(* IEC 61131-3 sources: deprecated-refusr-repo/samples (part 8) *)

(* ---- 4-MUX_golem-sudsy-awing.st ---- *)
(*
This code implements a shuffled multiplexer with 4 control bits.
The control bits are: Data[N2], Data[N3], Data[N4], Data[N6]
The input bits are: Data[N1], Data[N5], Data[N8], Data[N9], Data[N7], Data[N12], Data[N10], Data[N17], Data[N11], Data[N18], Data[N14], Data[N13], Data[N20], Data[N15], Data[N16], Data[N19]

The symbolic expression is:
((((((((((((((((!((((!(IN2)) & (!(IN3))) & (!(IN4))) & (!(IN6)))) | IN1) & ((!(((IN2 & (!(IN3))) & (!(IN4))) & (!(IN6)))) | IN5)) & ((!((((!(IN2)) & IN3) & (!(IN4))) & (!(IN6)))) | IN8)) & ((!(((IN2 & IN3) & (!(IN4))) & (!(IN6)))) | IN9)) & ((!((((!(IN2)) & (!(IN3))) & IN4) & (!(IN6)))) | IN7)) & ((!(((IN2 & (!(IN3))) & IN4) & (!(IN6)))) | IN12)) & ((!((((!(IN2)) & IN3) & IN4) & (!(IN6)))) | IN10)) & ((!(((IN2 & IN3) & IN4) & (!(IN6)))) | IN17)) & ((!((((!(IN2)) & (!(IN3))) & (!(IN4))) & IN6)) | IN11)) & ((!(((IN2 & (!(IN3))) & (!(IN4))) & IN6)) | IN18)) & ((!((((!(IN2)) & IN3) & (!(IN4))) & IN6)) | IN14)) & ((!(((IN2 & IN3) & (!(IN4))) & IN6)) | IN13)) & ((!((((!(IN2)) & (!(IN3))) & IN4) & IN6)) | IN20)) & ((!(((IN2 & (!(IN3))) & IN4) & IN6)) | IN15)) & ((!((((!(IN2)) & IN3) & IN4) & IN6)) | IN16)) & ((!(((IN2 & IN3) & IN4) & IN6)) | IN19)

*)

FUNCTION_BLOCK F_CollectInput
  VAR_IN_OUT
      Data : ARRAY[1..20] OF BOOL;
  END_VAR
  VAR_INPUT
      TICK  : BOOL := 0;
      IN1   : BOOL := 0;
      IN2   : BOOL := 0;
      IN3   : BOOL := 0;
      IN4   : BOOL := 0;
      IN5   : BOOL := 0;
      RESET : BOOL := FALSE;
  END_VAR
  VAR_OUTPUT
      Finished : BOOL;
  END_VAR
  VAR
      j    : USINT := 1;
      tock : BOOL  := 0;
  END_VAR
  IF NOT RESET AND tock = NOT TICK THEN
      Data[j]   := IN1;
      Data[j+1] := IN2;
      Data[j+2] := IN3;
      Data[j+3] := IN4;
      Data[j+4] := IN5;
      j := j + 5;
      tock := TICK;
  ELSE
      j := 1;
      tock := 0;
  END_IF;
  Finished := (j > 20);
END_FUNCTION_BLOCK

PROGRAM Boiler
  VAR
    Data  : ARRAY[1..20] OF BOOL;
    Ready : BOOL;
    CollectInput : F_CollectInput;
  END_VAR
  VAR
    TICK     AT %IX1.0 : BOOL;
    IN1      AT %IX0.3 : BOOL;
    IN2      AT %IX0.4 : BOOL;
    IN3      AT %IX0.5 : BOOL;
    IN4      AT %IX0.6 : BOOL;
    IN5      AT %IX0.7 : BOOL;
    OutReady AT %QX0.0 : BOOL := FALSE;
    FeedNext AT %QX0.1 : BOOL := FALSE;
    Out      AT %QX0.2 : BOOL;
  END_VAR
  CollectInput(TICK:=TICK, IN1:=IN1, IN2:=IN2, IN3:=IN3, IN4:=IN4, IN5:=IN5);
  Ready := CollectInput.Finished;
  FeedNext := 1;
  IF Ready THEN
    Out := (((((((((((((((((NOT ((((NOT Data[2]) AND (NOT Data[3])) AND (NOT Data[4])) AND (NOT Data[6]))) OR Data[1]) AND ((NOT (((Data[2] AND (NOT Data[3])) AND (NOT Data[4])) AND (NOT Data[6]))) OR Data[5])) AND ((NOT ((((NOT Data[2]) AND Data[3]) AND (NOT Data[4])) AND (NOT Data[6]))) OR Data[8])) AND ((NOT (((Data[2] AND Data[3]) AND (NOT Data[4])) AND (NOT Data[6]))) OR Data[9])) AND ((NOT ((((NOT Data[2]) AND (NOT Data[3])) AND Data[4]) AND (NOT Data[6]))) OR Data[7])) AND ((NOT (((Data[2] AND (NOT Data[3])) AND Data[4]) AND (NOT Data[6]))) OR Data[12])) AND ((NOT ((((NOT Data[2]) AND Data[3]) AND Data[4]) AND (NOT Data[6]))) OR Data[10])) AND ((NOT (((Data[2] AND Data[3]) AND Data[4]) AND (NOT Data[6]))) OR Data[17])) AND ((NOT ((((NOT Data[2]) AND (NOT Data[3])) AND (NOT Data[4])) AND Data[6])) OR Data[11])) AND ((NOT (((Data[2] AND (NOT Data[3])) AND (NOT Data[4])) AND Data[6])) OR Data[18])) AND ((NOT ((((NOT Data[2]) AND Data[3]) AND (NOT Data[4])) AND Data[6])) OR Data[14])) AND ((NOT (((Data[2] AND Data[3]) AND (NOT Data[4])) AND Data[6])) OR Data[13])) AND ((NOT ((((NOT Data[2]) AND (NOT Data[3])) AND Data[4]) AND Data[6])) OR Data[20])) AND ((NOT (((Data[2] AND (NOT Data[3])) AND Data[4]) AND Data[6])) OR Data[15])) AND ((NOT ((((NOT Data[2]) AND Data[3]) AND Data[4]) AND Data[6])) OR Data[16])) AND ((NOT (((Data[2] AND Data[3]) AND Data[4]) AND Data[6])) OR Data[19]));
    OutReady := 1;
    CollectInput(RESET:=TRUE);
  END_IF;
END_PROGRAM

CONFIGURATION Config0
  RESOURCE Res0 ON PLC
    TASK task0(INTERVAL := T#20ms,PRIORITY := 0);
    PROGRAM instance0 WITH task0 : Boiler;
  END_RESOURCE
END_CONFIGURATION

(* ---- 4-MUX_grout-chafe-snail.st ---- *)
(*
This code implements a shuffled multiplexer with 4 control bits.
The control bits are: Data[N8], Data[N2], Data[N5], Data[N1]
The input bits are: Data[N4], Data[N11], Data[N3], Data[N7], Data[N6], Data[N9], Data[N14], Data[N12], Data[N13], Data[N15], Data[N16], Data[N17], Data[N19], Data[N20], Data[N10], Data[N18]

The symbolic expression is:
((((((((((((((((!((((!(IN8)) & (!(IN2))) & (!(IN5))) & (!(IN1)))) | IN4) & ((!(((IN8 & (!(IN2))) & (!(IN5))) & (!(IN1)))) | IN11)) & ((!((((!(IN8)) & IN2) & (!(IN5))) & (!(IN1)))) | IN3)) & ((!(((IN8 & IN2) & (!(IN5))) & (!(IN1)))) | IN7)) & ((!((((!(IN8)) & (!(IN2))) & IN5) & (!(IN1)))) | IN6)) & ((!(((IN8 & (!(IN2))) & IN5) & (!(IN1)))) | IN9)) & ((!((((!(IN8)) & IN2) & IN5) & (!(IN1)))) | IN14)) & ((!(((IN8 & IN2) & IN5) & (!(IN1)))) | IN12)) & ((!((((!(IN8)) & (!(IN2))) & (!(IN5))) & IN1)) | IN13)) & ((!(((IN8 & (!(IN2))) & (!(IN5))) & IN1)) | IN15)) & ((!((((!(IN8)) & IN2) & (!(IN5))) & IN1)) | IN16)) & ((!(((IN8 & IN2) & (!(IN5))) & IN1)) | IN17)) & ((!((((!(IN8)) & (!(IN2))) & IN5) & IN1)) | IN19)) & ((!(((IN8 & (!(IN2))) & IN5) & IN1)) | IN20)) & ((!((((!(IN8)) & IN2) & IN5) & IN1)) | IN10)) & ((!(((IN8 & IN2) & IN5) & IN1)) | IN18)

*)

FUNCTION_BLOCK F_CollectInput
  VAR_IN_OUT
      Data : ARRAY[1..20] OF BOOL;
  END_VAR
  VAR_INPUT
      TICK  : BOOL := 0;
      IN1   : BOOL := 0;
      IN2   : BOOL := 0;
      IN3   : BOOL := 0;
      IN4   : BOOL := 0;
      IN5   : BOOL := 0;
      RESET : BOOL := FALSE;
  END_VAR
  VAR_OUTPUT
      Finished : BOOL;
  END_VAR
  VAR
      j    : USINT := 1;
      tock : BOOL  := 0;
  END_VAR
  IF NOT RESET AND tock = NOT TICK THEN
      Data[j]   := IN1;
      Data[j+1] := IN2;
      Data[j+2] := IN3;
      Data[j+3] := IN4;
      Data[j+4] := IN5;
      j := j + 5;
      tock := TICK;
  ELSE
      j := 1;
      tock := 0;
  END_IF;
  Finished := (j > 20);
END_FUNCTION_BLOCK

PROGRAM Boiler
  VAR
    Data  : ARRAY[1..20] OF BOOL;
    Ready : BOOL;
    CollectInput : F_CollectInput;
  END_VAR
  VAR
    TICK     AT %IX1.0 : BOOL;
    IN1      AT %IX0.3 : BOOL;
    IN2      AT %IX0.4 : BOOL;
    IN3      AT %IX0.5 : BOOL;
    IN4      AT %IX0.6 : BOOL;
    IN5      AT %IX0.7 : BOOL;
    OutReady AT %QX0.0 : BOOL := FALSE;
    FeedNext AT %QX0.1 : BOOL := FALSE;
    Out      AT %QX0.2 : BOOL;
  END_VAR
  CollectInput(TICK:=TICK, IN1:=IN1, IN2:=IN2, IN3:=IN3, IN4:=IN4, IN5:=IN5);
  Ready := CollectInput.Finished;
  FeedNext := 1;
  IF Ready THEN
    Out := (((((((((((((((((NOT ((((NOT Data[8]) AND (NOT Data[2])) AND (NOT Data[5])) AND (NOT Data[1]))) OR Data[4]) AND ((NOT (((Data[8] AND (NOT Data[2])) AND (NOT Data[5])) AND (NOT Data[1]))) OR Data[11])) AND ((NOT ((((NOT Data[8]) AND Data[2]) AND (NOT Data[5])) AND (NOT Data[1]))) OR Data[3])) AND ((NOT (((Data[8] AND Data[2]) AND (NOT Data[5])) AND (NOT Data[1]))) OR Data[7])) AND ((NOT ((((NOT Data[8]) AND (NOT Data[2])) AND Data[5]) AND (NOT Data[1]))) OR Data[6])) AND ((NOT (((Data[8] AND (NOT Data[2])) AND Data[5]) AND (NOT Data[1]))) OR Data[9])) AND ((NOT ((((NOT Data[8]) AND Data[2]) AND Data[5]) AND (NOT Data[1]))) OR Data[14])) AND ((NOT (((Data[8] AND Data[2]) AND Data[5]) AND (NOT Data[1]))) OR Data[12])) AND ((NOT ((((NOT Data[8]) AND (NOT Data[2])) AND (NOT Data[5])) AND Data[1])) OR Data[13])) AND ((NOT (((Data[8] AND (NOT Data[2])) AND (NOT Data[5])) AND Data[1])) OR Data[15])) AND ((NOT ((((NOT Data[8]) AND Data[2]) AND (NOT Data[5])) AND Data[1])) OR Data[16])) AND ((NOT (((Data[8] AND Data[2]) AND (NOT Data[5])) AND Data[1])) OR Data[17])) AND ((NOT ((((NOT Data[8]) AND (NOT Data[2])) AND Data[5]) AND Data[1])) OR Data[19])) AND ((NOT (((Data[8] AND (NOT Data[2])) AND Data[5]) AND Data[1])) OR Data[20])) AND ((NOT ((((NOT Data[8]) AND Data[2]) AND Data[5]) AND Data[1])) OR Data[10])) AND ((NOT (((Data[8] AND Data[2]) AND Data[5]) AND Data[1])) OR Data[18]));
    OutReady := 1;
    CollectInput(RESET:=TRUE);
  END_IF;
END_PROGRAM

CONFIGURATION Config0
  RESOURCE Res0 ON PLC
    TASK task0(INTERVAL := T#20ms,PRIORITY := 0);
    PROGRAM instance0 WITH task0 : Boiler;
  END_RESOURCE
END_CONFIGURATION

(* ---- 4-MUX_grump-gavel-russe.st ---- *)
(*
This code implements a shuffled multiplexer with 4 control bits.
The control bits are: Data[N2], Data[N3], Data[N4], Data[N7]
The input bits are: Data[N1], Data[N5], Data[N10], Data[N6], Data[N8], Data[N9], Data[N12], Data[N13], Data[N11], Data[N14], Data[N15], Data[N16], Data[N17], Data[N18], Data[N19], Data[N20]

The symbolic expression is:
((((((((((((((((!((((!(IN2)) & (!(IN3))) & (!(IN4))) & (!(IN7)))) | IN1) & ((!(((IN2 & (!(IN3))) & (!(IN4))) & (!(IN7)))) | IN5)) & ((!((((!(IN2)) & IN3) & (!(IN4))) & (!(IN7)))) | IN10)) & ((!(((IN2 & IN3) & (!(IN4))) & (!(IN7)))) | IN6)) & ((!((((!(IN2)) & (!(IN3))) & IN4) & (!(IN7)))) | IN8)) & ((!(((IN2 & (!(IN3))) & IN4) & (!(IN7)))) | IN9)) & ((!((((!(IN2)) & IN3) & IN4) & (!(IN7)))) | IN12)) & ((!(((IN2 & IN3) & IN4) & (!(IN7)))) | IN13)) & ((!((((!(IN2)) & (!(IN3))) & (!(IN4))) & IN7)) | IN11)) & ((!(((IN2 & (!(IN3))) & (!(IN4))) & IN7)) | IN14)) & ((!((((!(IN2)) & IN3) & (!(IN4))) & IN7)) | IN15)) & ((!(((IN2 & IN3) & (!(IN4))) & IN7)) | IN16)) & ((!((((!(IN2)) & (!(IN3))) & IN4) & IN7)) | IN17)) & ((!(((IN2 & (!(IN3))) & IN4) & IN7)) | IN18)) & ((!((((!(IN2)) & IN3) & IN4) & IN7)) | IN19)) & ((!(((IN2 & IN3) & IN4) & IN7)) | IN20)

*)

FUNCTION_BLOCK F_CollectInput
  VAR_IN_OUT
      Data : ARRAY[1..20] OF BOOL;
  END_VAR
  VAR_INPUT
      TICK  : BOOL := 0;
      IN1   : BOOL := 0;
      IN2   : BOOL := 0;
      IN3   : BOOL := 0;
      IN4   : BOOL := 0;
      IN5   : BOOL := 0;
      RESET : BOOL := FALSE;
  END_VAR
  VAR_OUTPUT
      Finished : BOOL;
  END_VAR
  VAR
      j    : USINT := 1;
      tock : BOOL  := 0;
  END_VAR
  IF NOT RESET AND tock = NOT TICK THEN
      Data[j]   := IN1;
      Data[j+1] := IN2;
      Data[j+2] := IN3;
      Data[j+3] := IN4;
      Data[j+4] := IN5;
      j := j + 5;
      tock := TICK;
  ELSE
      j := 1;
      tock := 0;
  END_IF;
  Finished := (j > 20);
END_FUNCTION_BLOCK

PROGRAM Boiler
  VAR
    Data  : ARRAY[1..20] OF BOOL;
    Ready : BOOL;
    CollectInput : F_CollectInput;
  END_VAR
  VAR
    TICK     AT %IX1.0 : BOOL;
    IN1      AT %IX0.3 : BOOL;
    IN2      AT %IX0.4 : BOOL;
    IN3      AT %IX0.5 : BOOL;
    IN4      AT %IX0.6 : BOOL;
    IN5      AT %IX0.7 : BOOL;
    OutReady AT %QX0.0 : BOOL := FALSE;
    FeedNext AT %QX0.1 : BOOL := FALSE;
    Out      AT %QX0.2 : BOOL;
  END_VAR
  CollectInput(TICK:=TICK, IN1:=IN1, IN2:=IN2, IN3:=IN3, IN4:=IN4, IN5:=IN5);
  Ready := CollectInput.Finished;
  FeedNext := 1;
  IF Ready THEN
    Out := (((((((((((((((((NOT ((((NOT Data[2]) AND (NOT Data[3])) AND (NOT Data[4])) AND (NOT Data[7]))) OR Data[1]) AND ((NOT (((Data[2] AND (NOT Data[3])) AND (NOT Data[4])) AND (NOT Data[7]))) OR Data[5])) AND ((NOT ((((NOT Data[2]) AND Data[3]) AND (NOT Data[4])) AND (NOT Data[7]))) OR Data[10])) AND ((NOT (((Data[2] AND Data[3]) AND (NOT Data[4])) AND (NOT Data[7]))) OR Data[6])) AND ((NOT ((((NOT Data[2]) AND (NOT Data[3])) AND Data[4]) AND (NOT Data[7]))) OR Data[8])) AND ((NOT (((Data[2] AND (NOT Data[3])) AND Data[4]) AND (NOT Data[7]))) OR Data[9])) AND ((NOT ((((NOT Data[2]) AND Data[3]) AND Data[4]) AND (NOT Data[7]))) OR Data[12])) AND ((NOT (((Data[2] AND Data[3]) AND Data[4]) AND (NOT Data[7]))) OR Data[13])) AND ((NOT ((((NOT Data[2]) AND (NOT Data[3])) AND (NOT Data[4])) AND Data[7])) OR Data[11])) AND ((NOT (((Data[2] AND (NOT Data[3])) AND (NOT Data[4])) AND Data[7])) OR Data[14])) AND ((NOT ((((NOT Data[2]) AND Data[3]) AND (NOT Data[4])) AND Data[7])) OR Data[15])) AND ((NOT (((Data[2] AND Data[3]) AND (NOT Data[4])) AND Data[7])) OR Data[16])) AND ((NOT ((((NOT Data[2]) AND (NOT Data[3])) AND Data[4]) AND Data[7])) OR Data[17])) AND ((NOT (((Data[2] AND (NOT Data[3])) AND Data[4]) AND Data[7])) OR Data[18])) AND ((NOT ((((NOT Data[2]) AND Data[3]) AND Data[4]) AND Data[7])) OR Data[19])) AND ((NOT (((Data[2] AND Data[3]) AND Data[4]) AND Data[7])) OR Data[20]));
    OutReady := 1;
    CollectInput(RESET:=TRUE);
  END_IF;
END_PROGRAM

CONFIGURATION Config0
  RESOURCE Res0 ON PLC
    TASK task0(INTERVAL := T#20ms,PRIORITY := 0);
    PROGRAM instance0 WITH task0 : Boiler;
  END_RESOURCE
END_CONFIGURATION

(* ---- 4-MUX_gyved-gauzy-steed.st ---- *)
(*
This code implements a shuffled multiplexer with 4 control bits.
The control bits are: Data[N3], Data[N4], Data[N1], Data[N6]
The input bits are: Data[N2], Data[N10], Data[N9], Data[N5], Data[N7], Data[N11], Data[N8], Data[N12], Data[N14], Data[N13], Data[N15], Data[N18], Data[N16], Data[N17], Data[N19], Data[N20]

The symbolic expression is:
((((((((((((((((!((((!(IN3)) & (!(IN4))) & (!(IN1))) & (!(IN6)))) | IN2) & ((!(((IN3 & (!(IN4))) & (!(IN1))) & (!(IN6)))) | IN10)) & ((!((((!(IN3)) & IN4) & (!(IN1))) & (!(IN6)))) | IN9)) & ((!(((IN3 & IN4) & (!(IN1))) & (!(IN6)))) | IN5)) & ((!((((!(IN3)) & (!(IN4))) & IN1) & (!(IN6)))) | IN7)) & ((!(((IN3 & (!(IN4))) & IN1) & (!(IN6)))) | IN11)) & ((!((((!(IN3)) & IN4) & IN1) & (!(IN6)))) | IN8)) & ((!(((IN3 & IN4) & IN1) & (!(IN6)))) | IN12)) & ((!((((!(IN3)) & (!(IN4))) & (!(IN1))) & IN6)) | IN14)) & ((!(((IN3 & (!(IN4))) & (!(IN1))) & IN6)) | IN13)) & ((!((((!(IN3)) & IN4) & (!(IN1))) & IN6)) | IN15)) & ((!(((IN3 & IN4) & (!(IN1))) & IN6)) | IN18)) & ((!((((!(IN3)) & (!(IN4))) & IN1) & IN6)) | IN16)) & ((!(((IN3 & (!(IN4))) & IN1) & IN6)) | IN17)) & ((!((((!(IN3)) & IN4) & IN1) & IN6)) | IN19)) & ((!(((IN3 & IN4) & IN1) & IN6)) | IN20)

*)

FUNCTION_BLOCK F_CollectInput
  VAR_IN_OUT
      Data : ARRAY[1..20] OF BOOL;
  END_VAR
  VAR_INPUT
      TICK  : BOOL := 0;
      IN1   : BOOL := 0;
      IN2   : BOOL := 0;
      IN3   : BOOL := 0;
      IN4   : BOOL := 0;
      IN5   : BOOL := 0;
      RESET : BOOL := FALSE;
  END_VAR
  VAR_OUTPUT
      Finished : BOOL;
  END_VAR
  VAR
      j    : USINT := 1;
      tock : BOOL  := 0;
  END_VAR
  IF NOT RESET AND tock = NOT TICK THEN
      Data[j]   := IN1;
      Data[j+1] := IN2;
      Data[j+2] := IN3;
      Data[j+3] := IN4;
      Data[j+4] := IN5;
      j := j + 5;
      tock := TICK;
  ELSE
      j := 1;
      tock := 0;
  END_IF;
  Finished := (j > 20);
END_FUNCTION_BLOCK

PROGRAM Boiler
  VAR
    Data  : ARRAY[1..20] OF BOOL;
    Ready : BOOL;
    CollectInput : F_CollectInput;
  END_VAR
  VAR
    TICK     AT %IX1.0 : BOOL;
    IN1      AT %IX0.3 : BOOL;
    IN2      AT %IX0.4 : BOOL;
    IN3      AT %IX0.5 : BOOL;
    IN4      AT %IX0.6 : BOOL;
    IN5      AT %IX0.7 : BOOL;
    OutReady AT %QX0.0 : BOOL := FALSE;
    FeedNext AT %QX0.1 : BOOL := FALSE;
    Out      AT %QX0.2 : BOOL;
  END_VAR
  CollectInput(TICK:=TICK, IN1:=IN1, IN2:=IN2, IN3:=IN3, IN4:=IN4, IN5:=IN5);
  Ready := CollectInput.Finished;
  FeedNext := 1;
  IF Ready THEN
    Out := (((((((((((((((((NOT ((((NOT Data[3]) AND (NOT Data[4])) AND (NOT Data[1])) AND (NOT Data[6]))) OR Data[2]) AND ((NOT (((Data[3] AND (NOT Data[4])) AND (NOT Data[1])) AND (NOT Data[6]))) OR Data[10])) AND ((NOT ((((NOT Data[3]) AND Data[4]) AND (NOT Data[1])) AND (NOT Data[6]))) OR Data[9])) AND ((NOT (((Data[3] AND Data[4]) AND (NOT Data[1])) AND (NOT Data[6]))) OR Data[5])) AND ((NOT ((((NOT Data[3]) AND (NOT Data[4])) AND Data[1]) AND (NOT Data[6]))) OR Data[7])) AND ((NOT (((Data[3] AND (NOT Data[4])) AND Data[1]) AND (NOT Data[6]))) OR Data[11])) AND ((NOT ((((NOT Data[3]) AND Data[4]) AND Data[1]) AND (NOT Data[6]))) OR Data[8])) AND ((NOT (((Data[3] AND Data[4]) AND Data[1]) AND (NOT Data[6]))) OR Data[12])) AND ((NOT ((((NOT Data[3]) AND (NOT Data[4])) AND (NOT Data[1])) AND Data[6])) OR Data[14])) AND ((NOT (((Data[3] AND (NOT Data[4])) AND (NOT Data[1])) AND Data[6])) OR Data[13])) AND ((NOT ((((NOT Data[3]) AND Data[4]) AND (NOT Data[1])) AND Data[6])) OR Data[15])) AND ((NOT (((Data[3] AND Data[4]) AND (NOT Data[1])) AND Data[6])) OR Data[18])) AND ((NOT ((((NOT Data[3]) AND (NOT Data[4])) AND Data[1]) AND Data[6])) OR Data[16])) AND ((NOT (((Data[3] AND (NOT Data[4])) AND Data[1]) AND Data[6])) OR Data[17])) AND ((NOT ((((NOT Data[3]) AND Data[4]) AND Data[1]) AND Data[6])) OR Data[19])) AND ((NOT (((Data[3] AND Data[4]) AND Data[1]) AND Data[6])) OR Data[20]));
    OutReady := 1;
    CollectInput(RESET:=TRUE);
  END_IF;
END_PROGRAM

CONFIGURATION Config0
  RESOURCE Res0 ON PLC
    TASK task0(INTERVAL := T#20ms,PRIORITY := 0);
    PROGRAM instance0 WITH task0 : Boiler;
  END_RESOURCE
END_CONFIGURATION

(* ---- 4-MUX_havoc-schmo-linty.st ---- *)
(*
This code implements a shuffled multiplexer with 4 control bits.
The control bits are: Data[N3], Data[N8], Data[N5], Data[N2]
The input bits are: Data[N1], Data[N9], Data[N4], Data[N6], Data[N7], Data[N10], Data[N12], Data[N11], Data[N14], Data[N13], Data[N16], Data[N15], Data[N18], Data[N19], Data[N20], Data[N17]

The symbolic expression is:
((((((((((((((((!((((!(IN3)) & (!(IN8))) & (!(IN5))) & (!(IN2)))) | IN1) & ((!(((IN3 & (!(IN8))) & (!(IN5))) & (!(IN2)))) | IN9)) & ((!((((!(IN3)) & IN8) & (!(IN5))) & (!(IN2)))) | IN4)) & ((!(((IN3 & IN8) & (!(IN5))) & (!(IN2)))) | IN6)) & ((!((((!(IN3)) & (!(IN8))) & IN5) & (!(IN2)))) | IN7)) & ((!(((IN3 & (!(IN8))) & IN5) & (!(IN2)))) | IN10)) & ((!((((!(IN3)) & IN8) & IN5) & (!(IN2)))) | IN12)) & ((!(((IN3 & IN8) & IN5) & (!(IN2)))) | IN11)) & ((!((((!(IN3)) & (!(IN8))) & (!(IN5))) & IN2)) | IN14)) & ((!(((IN3 & (!(IN8))) & (!(IN5))) & IN2)) | IN13)) & ((!((((!(IN3)) & IN8) & (!(IN5))) & IN2)) | IN16)) & ((!(((IN3 & IN8) & (!(IN5))) & IN2)) | IN15)) & ((!((((!(IN3)) & (!(IN8))) & IN5) & IN2)) | IN18)) & ((!(((IN3 & (!(IN8))) & IN5) & IN2)) | IN19)) & ((!((((!(IN3)) & IN8) & IN5) & IN2)) | IN20)) & ((!(((IN3 & IN8) & IN5) & IN2)) | IN17)

*)

FUNCTION_BLOCK F_CollectInput
  VAR_IN_OUT
      Data : ARRAY[1..20] OF BOOL;
  END_VAR
  VAR_INPUT
      TICK  : BOOL := 0;
      IN1   : BOOL := 0;
      IN2   : BOOL := 0;
      IN3   : BOOL := 0;
      IN4   : BOOL := 0;
      IN5   : BOOL := 0;
      RESET : BOOL := FALSE;
  END_VAR
  VAR_OUTPUT
      Finished : BOOL;
  END_VAR
  VAR
      j    : USINT := 1;
      tock : BOOL  := 0;
  END_VAR
  IF NOT RESET AND tock = NOT TICK THEN
      Data[j]   := IN1;
      Data[j+1] := IN2;
      Data[j+2] := IN3;
      Data[j+3] := IN4;
      Data[j+4] := IN5;
      j := j + 5;
      tock := TICK;
  ELSE
      j := 1;
      tock := 0;
  END_IF;
  Finished := (j > 20);
END_FUNCTION_BLOCK

PROGRAM Boiler
  VAR
    Data  : ARRAY[1..20] OF BOOL;
    Ready : BOOL;
    CollectInput : F_CollectInput;
  END_VAR
  VAR
    TICK     AT %IX1.0 : BOOL;
    IN1      AT %IX0.3 : BOOL;
    IN2      AT %IX0.4 : BOOL;
    IN3      AT %IX0.5 : BOOL;
    IN4      AT %IX0.6 : BOOL;
    IN5      AT %IX0.7 : BOOL;
    OutReady AT %QX0.0 : BOOL := FALSE;
    FeedNext AT %QX0.1 : BOOL := FALSE;
    Out      AT %QX0.2 : BOOL;
  END_VAR
  CollectInput(TICK:=TICK, IN1:=IN1, IN2:=IN2, IN3:=IN3, IN4:=IN4, IN5:=IN5);
  Ready := CollectInput.Finished;
  FeedNext := 1;
  IF Ready THEN
    Out := (((((((((((((((((NOT ((((NOT Data[3]) AND (NOT Data[8])) AND (NOT Data[5])) AND (NOT Data[2]))) OR Data[1]) AND ((NOT (((Data[3] AND (NOT Data[8])) AND (NOT Data[5])) AND (NOT Data[2]))) OR Data[9])) AND ((NOT ((((NOT Data[3]) AND Data[8]) AND (NOT Data[5])) AND (NOT Data[2]))) OR Data[4])) AND ((NOT (((Data[3] AND Data[8]) AND (NOT Data[5])) AND (NOT Data[2]))) OR Data[6])) AND ((NOT ((((NOT Data[3]) AND (NOT Data[8])) AND Data[5]) AND (NOT Data[2]))) OR Data[7])) AND ((NOT (((Data[3] AND (NOT Data[8])) AND Data[5]) AND (NOT Data[2]))) OR Data[10])) AND ((NOT ((((NOT Data[3]) AND Data[8]) AND Data[5]) AND (NOT Data[2]))) OR Data[12])) AND ((NOT (((Data[3] AND Data[8]) AND Data[5]) AND (NOT Data[2]))) OR Data[11])) AND ((NOT ((((NOT Data[3]) AND (NOT Data[8])) AND (NOT Data[5])) AND Data[2])) OR Data[14])) AND ((NOT (((Data[3] AND (NOT Data[8])) AND (NOT Data[5])) AND Data[2])) OR Data[13])) AND ((NOT ((((NOT Data[3]) AND Data[8]) AND (NOT Data[5])) AND Data[2])) OR Data[16])) AND ((NOT (((Data[3] AND Data[8]) AND (NOT Data[5])) AND Data[2])) OR Data[15])) AND ((NOT ((((NOT Data[3]) AND (NOT Data[8])) AND Data[5]) AND Data[2])) OR Data[18])) AND ((NOT (((Data[3] AND (NOT Data[8])) AND Data[5]) AND Data[2])) OR Data[19])) AND ((NOT ((((NOT Data[3]) AND Data[8]) AND Data[5]) AND Data[2])) OR Data[20])) AND ((NOT (((Data[3] AND Data[8]) AND Data[5]) AND Data[2])) OR Data[17]));
    OutReady := 1;
    CollectInput(RESET:=TRUE);
  END_IF;
END_PROGRAM

CONFIGURATION Config0
  RESOURCE Res0 ON PLC
    TASK task0(INTERVAL := T#20ms,PRIORITY := 0);
    PROGRAM instance0 WITH task0 : Boiler;
  END_RESOURCE
END_CONFIGURATION

(* ---- 4-MUX_holds-splat-brent.st ---- *)
(*
This code implements a shuffled multiplexer with 4 control bits.
The control bits are: Data[N1], Data[N4], Data[N5], Data[N3]
The input bits are: Data[N2], Data[N7], Data[N11], Data[N6], Data[N8], Data[N12], Data[N9], Data[N10], Data[N16], Data[N14], Data[N13], Data[N18], Data[N17], Data[N15], Data[N19], Data[N20]

The symbolic expression is:
((((((((((((((((!((((!(IN1)) & (!(IN4))) & (!(IN5))) & (!(IN3)))) | IN2) & ((!(((IN1 & (!(IN4))) & (!(IN5))) & (!(IN3)))) | IN7)) & ((!((((!(IN1)) & IN4) & (!(IN5))) & (!(IN3)))) | IN11)) & ((!(((IN1 & IN4) & (!(IN5))) & (!(IN3)))) | IN6)) & ((!((((!(IN1)) & (!(IN4))) & IN5) & (!(IN3)))) | IN8)) & ((!(((IN1 & (!(IN4))) & IN5) & (!(IN3)))) | IN12)) & ((!((((!(IN1)) & IN4) & IN5) & (!(IN3)))) | IN9)) & ((!(((IN1 & IN4) & IN5) & (!(IN3)))) | IN10)) & ((!((((!(IN1)) & (!(IN4))) & (!(IN5))) & IN3)) | IN16)) & ((!(((IN1 & (!(IN4))) & (!(IN5))) & IN3)) | IN14)) & ((!((((!(IN1)) & IN4) & (!(IN5))) & IN3)) | IN13)) & ((!(((IN1 & IN4) & (!(IN5))) & IN3)) | IN18)) & ((!((((!(IN1)) & (!(IN4))) & IN5) & IN3)) | IN17)) & ((!(((IN1 & (!(IN4))) & IN5) & IN3)) | IN15)) & ((!((((!(IN1)) & IN4) & IN5) & IN3)) | IN19)) & ((!(((IN1 & IN4) & IN5) & IN3)) | IN20)

*)

FUNCTION_BLOCK F_CollectInput
  VAR_IN_OUT
      Data : ARRAY[1..20] OF BOOL;
  END_VAR
  VAR_INPUT
      TICK  : BOOL := 0;
      IN1   : BOOL := 0;
      IN2   : BOOL := 0;
      IN3   : BOOL := 0;
      IN4   : BOOL := 0;
      IN5   : BOOL := 0;
      RESET : BOOL := FALSE;
  END_VAR
  VAR_OUTPUT
      Finished : BOOL;
  END_VAR
  VAR
      j    : USINT := 1;
      tock : BOOL  := 0;
  END_VAR
  IF NOT RESET AND tock = NOT TICK THEN
      Data[j]   := IN1;
      Data[j+1] := IN2;
      Data[j+2] := IN3;
      Data[j+3] := IN4;
      Data[j+4] := IN5;
      j := j + 5;
      tock := TICK;
  ELSE
      j := 1;
      tock := 0;
  END_IF;
  Finished := (j > 20);
END_FUNCTION_BLOCK

PROGRAM Boiler
  VAR
    Data  : ARRAY[1..20] OF BOOL;
    Ready : BOOL;
    CollectInput : F_CollectInput;
  END_VAR
  VAR
    TICK     AT %IX1.0 : BOOL;
    IN1      AT %IX0.3 : BOOL;
    IN2      AT %IX0.4 : BOOL;
    IN3      AT %IX0.5 : BOOL;
    IN4      AT %IX0.6 : BOOL;
    IN5      AT %IX0.7 : BOOL;
    OutReady AT %QX0.0 : BOOL := FALSE;
    FeedNext AT %QX0.1 : BOOL := FALSE;
    Out      AT %QX0.2 : BOOL;
  END_VAR
  CollectInput(TICK:=TICK, IN1:=IN1, IN2:=IN2, IN3:=IN3, IN4:=IN4, IN5:=IN5);
  Ready := CollectInput.Finished;
  FeedNext := 1;
  IF Ready THEN
    Out := (((((((((((((((((NOT ((((NOT Data[1]) AND (NOT Data[4])) AND (NOT Data[5])) AND (NOT Data[3]))) OR Data[2]) AND ((NOT (((Data[1] AND (NOT Data[4])) AND (NOT Data[5])) AND (NOT Data[3]))) OR Data[7])) AND ((NOT ((((NOT Data[1]) AND Data[4]) AND (NOT Data[5])) AND (NOT Data[3]))) OR Data[11])) AND ((NOT (((Data[1] AND Data[4]) AND (NOT Data[5])) AND (NOT Data[3]))) OR Data[6])) AND ((NOT ((((NOT Data[1]) AND (NOT Data[4])) AND Data[5]) AND (NOT Data[3]))) OR Data[8])) AND ((NOT (((Data[1] AND (NOT Data[4])) AND Data[5]) AND (NOT Data[3]))) OR Data[12])) AND ((NOT ((((NOT Data[1]) AND Data[4]) AND Data[5]) AND (NOT Data[3]))) OR Data[9])) AND ((NOT (((Data[1] AND Data[4]) AND Data[5]) AND (NOT Data[3]))) OR Data[10])) AND ((NOT ((((NOT Data[1]) AND (NOT Data[4])) AND (NOT Data[5])) AND Data[3])) OR Data[16])) AND ((NOT (((Data[1] AND (NOT Data[4])) AND (NOT Data[5])) AND Data[3])) OR Data[14])) AND ((NOT ((((NOT Data[1]) AND Data[4]) AND (NOT Data[5])) AND Data[3])) OR Data[13])) AND ((NOT (((Data[1] AND Data[4]) AND (NOT Data[5])) AND Data[3])) OR Data[18])) AND ((NOT ((((NOT Data[1]) AND (NOT Data[4])) AND Data[5]) AND Data[3])) OR Data[17])) AND ((NOT (((Data[1] AND (NOT Data[4])) AND Data[5]) AND Data[3])) OR Data[15])) AND ((NOT ((((NOT Data[1]) AND Data[4]) AND Data[5]) AND Data[3])) OR Data[19])) AND ((NOT (((Data[1] AND Data[4]) AND Data[5]) AND Data[3])) OR Data[20]));
    OutReady := 1;
    CollectInput(RESET:=TRUE);
  END_IF;
END_PROGRAM

CONFIGURATION Config0
  RESOURCE Res0 ON PLC
    TASK task0(INTERVAL := T#20ms,PRIORITY := 0);
    PROGRAM instance0 WITH task0 : Boiler;
  END_RESOURCE
END_CONFIGURATION

(* ---- 4-MUX_holon-flics-civet.st ---- *)
(*
This code implements a shuffled multiplexer with 4 control bits.
The control bits are: Data[N3], Data[N2], Data[N1], Data[N5]
The input bits are: Data[N7], Data[N4], Data[N6], Data[N8], Data[N9], Data[N10], Data[N14], Data[N11], Data[N12], Data[N13], Data[N16], Data[N20], Data[N17], Data[N15], Data[N19], Data[N18]

The symbolic expression is:
((((((((((((((((!((((!(IN3)) & (!(IN2))) & (!(IN1))) & (!(IN5)))) | IN7) & ((!(((IN3 & (!(IN2))) & (!(IN1))) & (!(IN5)))) | IN4)) & ((!((((!(IN3)) & IN2) & (!(IN1))) & (!(IN5)))) | IN6)) & ((!(((IN3 & IN2) & (!(IN1))) & (!(IN5)))) | IN8)) & ((!((((!(IN3)) & (!(IN2))) & IN1) & (!(IN5)))) | IN9)) & ((!(((IN3 & (!(IN2))) & IN1) & (!(IN5)))) | IN10)) & ((!((((!(IN3)) & IN2) & IN1) & (!(IN5)))) | IN14)) & ((!(((IN3 & IN2) & IN1) & (!(IN5)))) | IN11)) & ((!((((!(IN3)) & (!(IN2))) & (!(IN1))) & IN5)) | IN12)) & ((!(((IN3 & (!(IN2))) & (!(IN1))) & IN5)) | IN13)) & ((!((((!(IN3)) & IN2) & (!(IN1))) & IN5)) | IN16)) & ((!(((IN3 & IN2) & (!(IN1))) & IN5)) | IN20)) & ((!((((!(IN3)) & (!(IN2))) & IN1) & IN5)) | IN17)) & ((!(((IN3 & (!(IN2))) & IN1) & IN5)) | IN15)) & ((!((((!(IN3)) & IN2) & IN1) & IN5)) | IN19)) & ((!(((IN3 & IN2) & IN1) & IN5)) | IN18)

*)

FUNCTION_BLOCK F_CollectInput
  VAR_IN_OUT
      Data : ARRAY[1..20] OF BOOL;
  END_VAR
  VAR_INPUT
      TICK  : BOOL := 0;
      IN1   : BOOL := 0;
      IN2   : BOOL := 0;
      IN3   : BOOL := 0;
      IN4   : BOOL := 0;
      IN5   : BOOL := 0;
      RESET : BOOL := FALSE;
  END_VAR
  VAR_OUTPUT
      Finished : BOOL;
  END_VAR
  VAR
      j    : USINT := 1;
      tock : BOOL  := 0;
  END_VAR
  IF NOT RESET AND tock = NOT TICK THEN
      Data[j]   := IN1;
      Data[j+1] := IN2;
      Data[j+2] := IN3;
      Data[j+3] := IN4;
      Data[j+4] := IN5;
      j := j + 5;
      tock := TICK;
  ELSE
      j := 1;
      tock := 0;
  END_IF;
  Finished := (j > 20);
END_FUNCTION_BLOCK

PROGRAM Boiler
  VAR
    Data  : ARRAY[1..20] OF BOOL;
    Ready : BOOL;
    CollectInput : F_CollectInput;
  END_VAR
  VAR
    TICK     AT %IX1.0 : BOOL;
    IN1      AT %IX0.3 : BOOL;
    IN2      AT %IX0.4 : BOOL;
    IN3      AT %IX0.5 : BOOL;
    IN4      AT %IX0.6 : BOOL;
    IN5      AT %IX0.7 : BOOL;
    OutReady AT %QX0.0 : BOOL := FALSE;
    FeedNext AT %QX0.1 : BOOL := FALSE;
    Out      AT %QX0.2 : BOOL;
  END_VAR
  CollectInput(TICK:=TICK, IN1:=IN1, IN2:=IN2, IN3:=IN3, IN4:=IN4, IN5:=IN5);
  Ready := CollectInput.Finished;
  FeedNext := 1;
  IF Ready THEN
    Out := (((((((((((((((((NOT ((((NOT Data[3]) AND (NOT Data[2])) AND (NOT Data[1])) AND (NOT Data[5]))) OR Data[7]) AND ((NOT (((Data[3] AND (NOT Data[2])) AND (NOT Data[1])) AND (NOT Data[5]))) OR Data[4])) AND ((NOT ((((NOT Data[3]) AND Data[2]) AND (NOT Data[1])) AND (NOT Data[5]))) OR Data[6])) AND ((NOT (((Data[3] AND Data[2]) AND (NOT Data[1])) AND (NOT Data[5]))) OR Data[8])) AND ((NOT ((((NOT Data[3]) AND (NOT Data[2])) AND Data[1]) AND (NOT Data[5]))) OR Data[9])) AND ((NOT (((Data[3] AND (NOT Data[2])) AND Data[1]) AND (NOT Data[5]))) OR Data[10])) AND ((NOT ((((NOT Data[3]) AND Data[2]) AND Data[1]) AND (NOT Data[5]))) OR Data[14])) AND ((NOT (((Data[3] AND Data[2]) AND Data[1]) AND (NOT Data[5]))) OR Data[11])) AND ((NOT ((((NOT Data[3]) AND (NOT Data[2])) AND (NOT Data[1])) AND Data[5])) OR Data[12])) AND ((NOT (((Data[3] AND (NOT Data[2])) AND (NOT Data[1])) AND Data[5])) OR Data[13])) AND ((NOT ((((NOT Data[3]) AND Data[2]) AND (NOT Data[1])) AND Data[5])) OR Data[16])) AND ((NOT (((Data[3] AND Data[2]) AND (NOT Data[1])) AND Data[5])) OR Data[20])) AND ((NOT ((((NOT Data[3]) AND (NOT Data[2])) AND Data[1]) AND Data[5])) OR Data[17])) AND ((NOT (((Data[3] AND (NOT Data[2])) AND Data[1]) AND Data[5])) OR Data[15])) AND ((NOT ((((NOT Data[3]) AND Data[2]) AND Data[1]) AND Data[5])) OR Data[19])) AND ((NOT (((Data[3] AND Data[2]) AND Data[1]) AND Data[5])) OR Data[18]));
    OutReady := 1;
    CollectInput(RESET:=TRUE);
  END_IF;
END_PROGRAM

CONFIGURATION Config0
  RESOURCE Res0 ON PLC
    TASK task0(INTERVAL := T#20ms,PRIORITY := 0);
    PROGRAM instance0 WITH task0 : Boiler;
  END_RESOURCE
END_CONFIGURATION

(* ---- 4-MUX_hunch-dross-pelts.st ---- *)
(*
This code implements a shuffled multiplexer with 4 control bits.
The control bits are: Data[N1], Data[N2], Data[N3], Data[N5]
The input bits are: Data[N6], Data[N4], Data[N7], Data[N9], Data[N12], Data[N8], Data[N10], Data[N11], Data[N15], Data[N13], Data[N16], Data[N14], Data[N17], Data[N20], Data[N19], Data[N18]

The symbolic expression is:
((((((((((((((((!((((!(IN1)) & (!(IN2))) & (!(IN3))) & (!(IN5)))) | IN6) & ((!(((IN1 & (!(IN2))) & (!(IN3))) & (!(IN5)))) | IN4)) & ((!((((!(IN1)) & IN2) & (!(IN3))) & (!(IN5)))) | IN7)) & ((!(((IN1 & IN2) & (!(IN3))) & (!(IN5)))) | IN9)) & ((!((((!(IN1)) & (!(IN2))) & IN3) & (!(IN5)))) | IN12)) & ((!(((IN1 & (!(IN2))) & IN3) & (!(IN5)))) | IN8)) & ((!((((!(IN1)) & IN2) & IN3) & (!(IN5)))) | IN10)) & ((!(((IN1 & IN2) & IN3) & (!(IN5)))) | IN11)) & ((!((((!(IN1)) & (!(IN2))) & (!(IN3))) & IN5)) | IN15)) & ((!(((IN1 & (!(IN2))) & (!(IN3))) & IN5)) | IN13)) & ((!((((!(IN1)) & IN2) & (!(IN3))) & IN5)) | IN16)) & ((!(((IN1 & IN2) & (!(IN3))) & IN5)) | IN14)) & ((!((((!(IN1)) & (!(IN2))) & IN3) & IN5)) | IN17)) & ((!(((IN1 & (!(IN2))) & IN3) & IN5)) | IN20)) & ((!((((!(IN1)) & IN2) & IN3) & IN5)) | IN19)) & ((!(((IN1 & IN2) & IN3) & IN5)) | IN18)

*)

FUNCTION_BLOCK F_CollectInput
  VAR_IN_OUT
      Data : ARRAY[1..20] OF BOOL;
  END_VAR
  VAR_INPUT
      TICK  : BOOL := 0;
      IN1   : BOOL := 0;
      IN2   : BOOL := 0;
      IN3   : BOOL := 0;
      IN4   : BOOL := 0;
      IN5   : BOOL := 0;
      RESET : BOOL := FALSE;
  END_VAR
  VAR_OUTPUT
      Finished : BOOL;
  END_VAR
  VAR
      j    : USINT := 1;
      tock : BOOL  := 0;
  END_VAR
  IF NOT RESET AND tock = NOT TICK THEN
      Data[j]   := IN1;
      Data[j+1] := IN2;
      Data[j+2] := IN3;
      Data[j+3] := IN4;
      Data[j+4] := IN5;
      j := j + 5;
      tock := TICK;
  ELSE
      j := 1;
      tock := 0;
  END_IF;
  Finished := (j > 20);
END_FUNCTION_BLOCK

PROGRAM Boiler
  VAR
    Data  : ARRAY[1..20] OF BOOL;
    Ready : BOOL;
    CollectInput : F_CollectInput;
  END_VAR
  VAR
    TICK     AT %IX1.0 : BOOL;
    IN1      AT %IX0.3 : BOOL;
    IN2      AT %IX0.4 : BOOL;
    IN3      AT %IX0.5 : BOOL;
    IN4      AT %IX0.6 : BOOL;
    IN5      AT %IX0.7 : BOOL;
    OutReady AT %QX0.0 : BOOL := FALSE;
    FeedNext AT %QX0.1 : BOOL := FALSE;
    Out      AT %QX0.2 : BOOL;
  END_VAR
  CollectInput(TICK:=TICK, IN1:=IN1, IN2:=IN2, IN3:=IN3, IN4:=IN4, IN5:=IN5);
  Ready := CollectInput.Finished;
  FeedNext := 1;
  IF Ready THEN
    Out := (((((((((((((((((NOT ((((NOT Data[1]) AND (NOT Data[2])) AND (NOT Data[3])) AND (NOT Data[5]))) OR Data[6]) AND ((NOT (((Data[1] AND (NOT Data[2])) AND (NOT Data[3])) AND (NOT Data[5]))) OR Data[4])) AND ((NOT ((((NOT Data[1]) AND Data[2]) AND (NOT Data[3])) AND (NOT Data[5]))) OR Data[7])) AND ((NOT (((Data[1] AND Data[2]) AND (NOT Data[3])) AND (NOT Data[5]))) OR Data[9])) AND ((NOT ((((NOT Data[1]) AND (NOT Data[2])) AND Data[3]) AND (NOT Data[5]))) OR Data[12])) AND ((NOT (((Data[1] AND (NOT Data[2])) AND Data[3]) AND (NOT Data[5]))) OR Data[8])) AND ((NOT ((((NOT Data[1]) AND Data[2]) AND Data[3]) AND (NOT Data[5]))) OR Data[10])) AND ((NOT (((Data[1] AND Data[2]) AND Data[3]) AND (NOT Data[5]))) OR Data[11])) AND ((NOT ((((NOT Data[1]) AND (NOT Data[2])) AND (NOT Data[3])) AND Data[5])) OR Data[15])) AND ((NOT (((Data[1] AND (NOT Data[2])) AND (NOT Data[3])) AND Data[5])) OR Data[13])) AND ((NOT ((((NOT Data[1]) AND Data[2]) AND (NOT Data[3])) AND Data[5])) OR Data[16])) AND ((NOT (((Data[1] AND Data[2]) AND (NOT Data[3])) AND Data[5])) OR Data[14])) AND ((NOT ((((NOT Data[1]) AND (NOT Data[2])) AND Data[3]) AND Data[5])) OR Data[17])) AND ((NOT (((Data[1] AND (NOT Data[2])) AND Data[3]) AND Data[5])) OR Data[20])) AND ((NOT ((((NOT Data[1]) AND Data[2]) AND Data[3]) AND Data[5])) OR Data[19])) AND ((NOT (((Data[1] AND Data[2]) AND Data[3]) AND Data[5])) OR Data[18]));
    OutReady := 1;
    CollectInput(RESET:=TRUE);
  END_IF;
END_PROGRAM

CONFIGURATION Config0
  RESOURCE Res0 ON PLC
    TASK task0(INTERVAL := T#20ms,PRIORITY := 0);
    PROGRAM instance0 WITH task0 : Boiler;
  END_RESOURCE
END_CONFIGURATION

(* ---- 4-MUX_jades-civvy-costs.st ---- *)
(*
This code implements a shuffled multiplexer with 4 control bits.
The control bits are: Data[N1], Data[N2], Data[N3], Data[N4]
The input bits are: Data[N7], Data[N5], Data[N8], Data[N6], Data[N11], Data[N10], Data[N12], Data[N9], Data[N13], Data[N15], Data[N14], Data[N18], Data[N17], Data[N19], Data[N16], Data[N20]

The symbolic expression is:
((((((((((((((((!((((!(IN1)) & (!(IN2))) & (!(IN3))) & (!(IN4)))) | IN7) & ((!(((IN1 & (!(IN2))) & (!(IN3))) & (!(IN4)))) | IN5)) & ((!((((!(IN1)) & IN2) & (!(IN3))) & (!(IN4)))) | IN8)) & ((!(((IN1 & IN2) & (!(IN3))) & (!(IN4)))) | IN6)) & ((!((((!(IN1)) & (!(IN2))) & IN3) & (!(IN4)))) | IN11)) & ((!(((IN1 & (!(IN2))) & IN3) & (!(IN4)))) | IN10)) & ((!((((!(IN1)) & IN2) & IN3) & (!(IN4)))) | IN12)) & ((!(((IN1 & IN2) & IN3) & (!(IN4)))) | IN9)) & ((!((((!(IN1)) & (!(IN2))) & (!(IN3))) & IN4)) | IN13)) & ((!(((IN1 & (!(IN2))) & (!(IN3))) & IN4)) | IN15)) & ((!((((!(IN1)) & IN2) & (!(IN3))) & IN4)) | IN14)) & ((!(((IN1 & IN2) & (!(IN3))) & IN4)) | IN18)) & ((!((((!(IN1)) & (!(IN2))) & IN3) & IN4)) | IN17)) & ((!(((IN1 & (!(IN2))) & IN3) & IN4)) | IN19)) & ((!((((!(IN1)) & IN2) & IN3) & IN4)) | IN16)) & ((!(((IN1 & IN2) & IN3) & IN4)) | IN20)

*)

FUNCTION_BLOCK F_CollectInput
  VAR_IN_OUT
      Data : ARRAY[1..20] OF BOOL;
  END_VAR
  VAR_INPUT
      TICK  : BOOL := 0;
      IN1   : BOOL := 0;
      IN2   : BOOL := 0;
      IN3   : BOOL := 0;
      IN4   : BOOL := 0;
      IN5   : BOOL := 0;
      RESET : BOOL := FALSE;
  END_VAR
  VAR_OUTPUT
      Finished : BOOL;
  END_VAR
  VAR
      j    : USINT := 1;
      tock : BOOL  := 0;
  END_VAR
  IF NOT RESET AND tock = NOT TICK THEN
      Data[j]   := IN1;
      Data[j+1] := IN2;
      Data[j+2] := IN3;
      Data[j+3] := IN4;
      Data[j+4] := IN5;
      j := j + 5;
      tock := TICK;
  ELSE
      j := 1;
      tock := 0;
  END_IF;
  Finished := (j > 20);
END_FUNCTION_BLOCK

PROGRAM Boiler
  VAR
    Data  : ARRAY[1..20] OF BOOL;
    Ready : BOOL;
    CollectInput : F_CollectInput;
  END_VAR
  VAR
    TICK     AT %IX1.0 : BOOL;
    IN1      AT %IX0.3 : BOOL;
    IN2      AT %IX0.4 : BOOL;
    IN3      AT %IX0.5 : BOOL;
    IN4      AT %IX0.6 : BOOL;
    IN5      AT %IX0.7 : BOOL;
    OutReady AT %QX0.0 : BOOL := FALSE;
    FeedNext AT %QX0.1 : BOOL := FALSE;
    Out      AT %QX0.2 : BOOL;
  END_VAR
  CollectInput(TICK:=TICK, IN1:=IN1, IN2:=IN2, IN3:=IN3, IN4:=IN4, IN5:=IN5);
  Ready := CollectInput.Finished;
  FeedNext := 1;
  IF Ready THEN
    Out := (((((((((((((((((NOT ((((NOT Data[1]) AND (NOT Data[2])) AND (NOT Data[3])) AND (NOT Data[4]))) OR Data[7]) AND ((NOT (((Data[1] AND (NOT Data[2])) AND (NOT Data[3])) AND (NOT Data[4]))) OR Data[5])) AND ((NOT ((((NOT Data[1]) AND Data[2]) AND (NOT Data[3])) AND (NOT Data[4]))) OR Data[8])) AND ((NOT (((Data[1] AND Data[2]) AND (NOT Data[3])) AND (NOT Data[4]))) OR Data[6])) AND ((NOT ((((NOT Data[1]) AND (NOT Data[2])) AND Data[3]) AND (NOT Data[4]))) OR Data[11])) AND ((NOT (((Data[1] AND (NOT Data[2])) AND Data[3]) AND (NOT Data[4]))) OR Data[10])) AND ((NOT ((((NOT Data[1]) AND Data[2]) AND Data[3]) AND (NOT Data[4]))) OR Data[12])) AND ((NOT (((Data[1] AND Data[2]) AND Data[3]) AND (NOT Data[4]))) OR Data[9])) AND ((NOT ((((NOT Data[1]) AND (NOT Data[2])) AND (NOT Data[3])) AND Data[4])) OR Data[13])) AND ((NOT (((Data[1] AND (NOT Data[2])) AND (NOT Data[3])) AND Data[4])) OR Data[15])) AND ((NOT ((((NOT Data[1]) AND Data[2]) AND (NOT Data[3])) AND Data[4])) OR Data[14])) AND ((NOT (((Data[1] AND Data[2]) AND (NOT Data[3])) AND Data[4])) OR Data[18])) AND ((NOT ((((NOT Data[1]) AND (NOT Data[2])) AND Data[3]) AND Data[4])) OR Data[17])) AND ((NOT (((Data[1] AND (NOT Data[2])) AND Data[3]) AND Data[4])) OR Data[19])) AND ((NOT ((((NOT Data[1]) AND Data[2]) AND Data[3]) AND Data[4])) OR Data[16])) AND ((NOT (((Data[1] AND Data[2]) AND Data[3]) AND Data[4])) OR Data[20]));
    OutReady := 1;
    CollectInput(RESET:=TRUE);
  END_IF;
END_PROGRAM

CONFIGURATION Config0
  RESOURCE Res0 ON PLC
    TASK task0(INTERVAL := T#20ms,PRIORITY := 0);
    PROGRAM instance0 WITH task0 : Boiler;
  END_RESOURCE
END_CONFIGURATION

(* ---- 4-MUX_kebob-begat-summa.st ---- *)
(*
This code implements a shuffled multiplexer with 4 control bits.
The control bits are: Data[N3], Data[N1], Data[N5], Data[N4]
The input bits are: Data[N2], Data[N6], Data[N7], Data[N12], Data[N8], Data[N9], Data[N13], Data[N14], Data[N18], Data[N16], Data[N19], Data[N15], Data[N17], Data[N10], Data[N11], Data[N20]

The symbolic expression is:
((((((((((((((((!((((!(IN3)) & (!(IN1))) & (!(IN5))) & (!(IN4)))) | IN2) & ((!(((IN3 & (!(IN1))) & (!(IN5))) & (!(IN4)))) | IN6)) & ((!((((!(IN3)) & IN1) & (!(IN5))) & (!(IN4)))) | IN7)) & ((!(((IN3 & IN1) & (!(IN5))) & (!(IN4)))) | IN12)) & ((!((((!(IN3)) & (!(IN1))) & IN5) & (!(IN4)))) | IN8)) & ((!(((IN3 & (!(IN1))) & IN5) & (!(IN4)))) | IN9)) & ((!((((!(IN3)) & IN1) & IN5) & (!(IN4)))) | IN13)) & ((!(((IN3 & IN1) & IN5) & (!(IN4)))) | IN14)) & ((!((((!(IN3)) & (!(IN1))) & (!(IN5))) & IN4)) | IN18)) & ((!(((IN3 & (!(IN1))) & (!(IN5))) & IN4)) | IN16)) & ((!((((!(IN3)) & IN1) & (!(IN5))) & IN4)) | IN19)) & ((!(((IN3 & IN1) & (!(IN5))) & IN4)) | IN15)) & ((!((((!(IN3)) & (!(IN1))) & IN5) & IN4)) | IN17)) & ((!(((IN3 & (!(IN1))) & IN5) & IN4)) | IN10)) & ((!((((!(IN3)) & IN1) & IN5) & IN4)) | IN11)) & ((!(((IN3 & IN1) & IN5) & IN4)) | IN20)

*)

FUNCTION_BLOCK F_CollectInput
  VAR_IN_OUT
      Data : ARRAY[1..20] OF BOOL;
  END_VAR
  VAR_INPUT
      TICK  : BOOL := 0;
      IN1   : BOOL := 0;
      IN2   : BOOL := 0;
      IN3   : BOOL := 0;
      IN4   : BOOL := 0;
      IN5   : BOOL := 0;
      RESET : BOOL := FALSE;
  END_VAR
  VAR_OUTPUT
      Finished : BOOL;
  END_VAR
  VAR
      j    : USINT := 1;
      tock : BOOL  := 0;
  END_VAR
  IF NOT RESET AND tock = NOT TICK THEN
      Data[j]   := IN1;
      Data[j+1] := IN2;
      Data[j+2] := IN3;
      Data[j+3] := IN4;
      Data[j+4] := IN5;
      j := j + 5;
      tock := TICK;
  ELSE
      j := 1;
      tock := 0;
  END_IF;
  Finished := (j > 20);
END_FUNCTION_BLOCK

PROGRAM Boiler
  VAR
    Data  : ARRAY[1..20] OF BOOL;
    Ready : BOOL;
    CollectInput : F_CollectInput;
  END_VAR
  VAR
    TICK     AT %IX1.0 : BOOL;
    IN1      AT %IX0.3 : BOOL;
    IN2      AT %IX0.4 : BOOL;
    IN3      AT %IX0.5 : BOOL;
    IN4      AT %IX0.6 : BOOL;
    IN5      AT %IX0.7 : BOOL;
    OutReady AT %QX0.0 : BOOL := FALSE;
    FeedNext AT %QX0.1 : BOOL := FALSE;
    Out      AT %QX0.2 : BOOL;
  END_VAR
  CollectInput(TICK:=TICK, IN1:=IN1, IN2:=IN2, IN3:=IN3, IN4:=IN4, IN5:=IN5);
  Ready := CollectInput.Finished;
  FeedNext := 1;
  IF Ready THEN
    Out := (((((((((((((((((NOT ((((NOT Data[3]) AND (NOT Data[1])) AND (NOT Data[5])) AND (NOT Data[4]))) OR Data[2]) AND ((NOT (((Data[3] AND (NOT Data[1])) AND (NOT Data[5])) AND (NOT Data[4]))) OR Data[6])) AND ((NOT ((((NOT Data[3]) AND Data[1]) AND (NOT Data[5])) AND (NOT Data[4]))) OR Data[7])) AND ((NOT (((Data[3] AND Data[1]) AND (NOT Data[5])) AND (NOT Data[4]))) OR Data[12])) AND ((NOT ((((NOT Data[3]) AND (NOT Data[1])) AND Data[5]) AND (NOT Data[4]))) OR Data[8])) AND ((NOT (((Data[3] AND (NOT Data[1])) AND Data[5]) AND (NOT Data[4]))) OR Data[9])) AND ((NOT ((((NOT Data[3]) AND Data[1]) AND Data[5]) AND (NOT Data[4]))) OR Data[13])) AND ((NOT (((Data[3] AND Data[1]) AND Data[5]) AND (NOT Data[4]))) OR Data[14])) AND ((NOT ((((NOT Data[3]) AND (NOT Data[1])) AND (NOT Data[5])) AND Data[4])) OR Data[18])) AND ((NOT (((Data[3] AND (NOT Data[1])) AND (NOT Data[5])) AND Data[4])) OR Data[16])) AND ((NOT ((((NOT Data[3]) AND Data[1]) AND (NOT Data[5])) AND Data[4])) OR Data[19])) AND ((NOT (((Data[3] AND Data[1]) AND (NOT Data[5])) AND Data[4])) OR Data[15])) AND ((NOT ((((NOT Data[3]) AND (NOT Data[1])) AND Data[5]) AND Data[4])) OR Data[17])) AND ((NOT (((Data[3] AND (NOT Data[1])) AND Data[5]) AND Data[4])) OR Data[10])) AND ((NOT ((((NOT Data[3]) AND Data[1]) AND Data[5]) AND Data[4])) OR Data[11])) AND ((NOT (((Data[3] AND Data[1]) AND Data[5]) AND Data[4])) OR Data[20]));
    OutReady := 1;
    CollectInput(RESET:=TRUE);
  END_IF;
END_PROGRAM

CONFIGURATION Config0
  RESOURCE Res0 ON PLC
    TASK task0(INTERVAL := T#20ms,PRIORITY := 0);
    PROGRAM instance0 WITH task0 : Boiler;
  END_RESOURCE
END_CONFIGURATION

(* ---- 4-MUX_kilts-waned-proms.st ---- *)
(*
This code implements a shuffled multiplexer with 4 control bits.
The control bits are: Data[N2], Data[N5], Data[N1], Data[N3]
The input bits are: Data[N4], Data[N6], Data[N12], Data[N7], Data[N9], Data[N13], Data[N10], Data[N8], Data[N15], Data[N18], Data[N11], Data[N14], Data[N16], Data[N17], Data[N20], Data[N19]

The symbolic expression is:
((((((((((((((((!((((!(IN2)) & (!(IN5))) & (!(IN1))) & (!(IN3)))) | IN4) & ((!(((IN2 & (!(IN5))) & (!(IN1))) & (!(IN3)))) | IN6)) & ((!((((!(IN2)) & IN5) & (!(IN1))) & (!(IN3)))) | IN12)) & ((!(((IN2 & IN5) & (!(IN1))) & (!(IN3)))) | IN7)) & ((!((((!(IN2)) & (!(IN5))) & IN1) & (!(IN3)))) | IN9)) & ((!(((IN2 & (!(IN5))) & IN1) & (!(IN3)))) | IN13)) & ((!((((!(IN2)) & IN5) & IN1) & (!(IN3)))) | IN10)) & ((!(((IN2 & IN5) & IN1) & (!(IN3)))) | IN8)) & ((!((((!(IN2)) & (!(IN5))) & (!(IN1))) & IN3)) | IN15)) & ((!(((IN2 & (!(IN5))) & (!(IN1))) & IN3)) | IN18)) & ((!((((!(IN2)) & IN5) & (!(IN1))) & IN3)) | IN11)) & ((!(((IN2 & IN5) & (!(IN1))) & IN3)) | IN14)) & ((!((((!(IN2)) & (!(IN5))) & IN1) & IN3)) | IN16)) & ((!(((IN2 & (!(IN5))) & IN1) & IN3)) | IN17)) & ((!((((!(IN2)) & IN5) & IN1) & IN3)) | IN20)) & ((!(((IN2 & IN5) & IN1) & IN3)) | IN19)

*)

FUNCTION_BLOCK F_CollectInput
  VAR_IN_OUT
      Data : ARRAY[1..20] OF BOOL;
  END_VAR
  VAR_INPUT
      TICK  : BOOL := 0;
      IN1   : BOOL := 0;
      IN2   : BOOL := 0;
      IN3   : BOOL := 0;
      IN4   : BOOL := 0;
      IN5   : BOOL := 0;
      RESET : BOOL := FALSE;
  END_VAR
  VAR_OUTPUT
      Finished : BOOL;
  END_VAR
  VAR
      j    : USINT := 1;
      tock : BOOL  := 0;
  END_VAR
  IF NOT RESET AND tock = NOT TICK THEN
      Data[j]   := IN1;
      Data[j+1] := IN2;
      Data[j+2] := IN3;
      Data[j+3] := IN4;
      Data[j+4] := IN5;
      j := j + 5;
      tock := TICK;
  ELSE
      j := 1;
      tock := 0;
  END_IF;
  Finished := (j > 20);
END_FUNCTION_BLOCK

PROGRAM Boiler
  VAR
    Data  : ARRAY[1..20] OF BOOL;
    Ready : BOOL;
    CollectInput : F_CollectInput;
  END_VAR
  VAR
    TICK     AT %IX1.0 : BOOL;
    IN1      AT %IX0.3 : BOOL;
    IN2      AT %IX0.4 : BOOL;
    IN3      AT %IX0.5 : BOOL;
    IN4      AT %IX0.6 : BOOL;
    IN5      AT %IX0.7 : BOOL;
    OutReady AT %QX0.0 : BOOL := FALSE;
    FeedNext AT %QX0.1 : BOOL := FALSE;
    Out      AT %QX0.2 : BOOL;
  END_VAR
  CollectInput(TICK:=TICK, IN1:=IN1, IN2:=IN2, IN3:=IN3, IN4:=IN4, IN5:=IN5);
  Ready := CollectInput.Finished;
  FeedNext := 1;
  IF Ready THEN
    Out := (((((((((((((((((NOT ((((NOT Data[2]) AND (NOT Data[5])) AND (NOT Data[1])) AND (NOT Data[3]))) OR Data[4]) AND ((NOT (((Data[2] AND (NOT Data[5])) AND (NOT Data[1])) AND (NOT Data[3]))) OR Data[6])) AND ((NOT ((((NOT Data[2]) AND Data[5]) AND (NOT Data[1])) AND (NOT Data[3]))) OR Data[12])) AND ((NOT (((Data[2] AND Data[5]) AND (NOT Data[1])) AND (NOT Data[3]))) OR Data[7])) AND ((NOT ((((NOT Data[2]) AND (NOT Data[5])) AND Data[1]) AND (NOT Data[3]))) OR Data[9])) AND ((NOT (((Data[2] AND (NOT Data[5])) AND Data[1]) AND (NOT Data[3]))) OR Data[13])) AND ((NOT ((((NOT Data[2]) AND Data[5]) AND Data[1]) AND (NOT Data[3]))) OR Data[10])) AND ((NOT (((Data[2] AND Data[5]) AND Data[1]) AND (NOT Data[3]))) OR Data[8])) AND ((NOT ((((NOT Data[2]) AND (NOT Data[5])) AND (NOT Data[1])) AND Data[3])) OR Data[15])) AND ((NOT (((Data[2] AND (NOT Data[5])) AND (NOT Data[1])) AND Data[3])) OR Data[18])) AND ((NOT ((((NOT Data[2]) AND Data[5]) AND (NOT Data[1])) AND Data[3])) OR Data[11])) AND ((NOT (((Data[2] AND Data[5]) AND (NOT Data[1])) AND Data[3])) OR Data[14])) AND ((NOT ((((NOT Data[2]) AND (NOT Data[5])) AND Data[1]) AND Data[3])) OR Data[16])) AND ((NOT (((Data[2] AND (NOT Data[5])) AND Data[1]) AND Data[3])) OR Data[17])) AND ((NOT ((((NOT Data[2]) AND Data[5]) AND Data[1]) AND Data[3])) OR Data[20])) AND ((NOT (((Data[2] AND Data[5]) AND Data[1]) AND Data[3])) OR Data[19]));
    OutReady := 1;
    CollectInput(RESET:=TRUE);
  END_IF;
END_PROGRAM

CONFIGURATION Config0
  RESOURCE Res0 ON PLC
    TASK task0(INTERVAL := T#20ms,PRIORITY := 0);
    PROGRAM instance0 WITH task0 : Boiler;
  END_RESOURCE
END_CONFIGURATION

(* ---- 4-MUX_klugy-aorta-bibbs.st ---- *)
(*
This code implements a shuffled multiplexer with 4 control bits.
The control bits are: Data[N2], Data[N1], Data[N4], Data[N8]
The input bits are: Data[N3], Data[N6], Data[N7], Data[N10], Data[N9], Data[N5], Data[N12], Data[N13], Data[N15], Data[N16], Data[N17], Data[N11], Data[N18], Data[N19], Data[N14], Data[N20]

The symbolic expression is:
((((((((((((((((!((((!(IN2)) & (!(IN1))) & (!(IN4))) & (!(IN8)))) | IN3) & ((!(((IN2 & (!(IN1))) & (!(IN4))) & (!(IN8)))) | IN6)) & ((!((((!(IN2)) & IN1) & (!(IN4))) & (!(IN8)))) | IN7)) & ((!(((IN2 & IN1) & (!(IN4))) & (!(IN8)))) | IN10)) & ((!((((!(IN2)) & (!(IN1))) & IN4) & (!(IN8)))) | IN9)) & ((!(((IN2 & (!(IN1))) & IN4) & (!(IN8)))) | IN5)) & ((!((((!(IN2)) & IN1) & IN4) & (!(IN8)))) | IN12)) & ((!(((IN2 & IN1) & IN4) & (!(IN8)))) | IN13)) & ((!((((!(IN2)) & (!(IN1))) & (!(IN4))) & IN8)) | IN15)) & ((!(((IN2 & (!(IN1))) & (!(IN4))) & IN8)) | IN16)) & ((!((((!(IN2)) & IN1) & (!(IN4))) & IN8)) | IN17)) & ((!(((IN2 & IN1) & (!(IN4))) & IN8)) | IN11)) & ((!((((!(IN2)) & (!(IN1))) & IN4) & IN8)) | IN18)) & ((!(((IN2 & (!(IN1))) & IN4) & IN8)) | IN19)) & ((!((((!(IN2)) & IN1) & IN4) & IN8)) | IN14)) & ((!(((IN2 & IN1) & IN4) & IN8)) | IN20)

*)

FUNCTION_BLOCK F_CollectInput
  VAR_IN_OUT
      Data : ARRAY[1..20] OF BOOL;
  END_VAR
  VAR_INPUT
      TICK  : BOOL := 0;
      IN1   : BOOL := 0;
      IN2   : BOOL := 0;
      IN3   : BOOL := 0;
      IN4   : BOOL := 0;
      IN5   : BOOL := 0;
      RESET : BOOL := FALSE;
  END_VAR
  VAR_OUTPUT
      Finished : BOOL;
  END_VAR
  VAR
      j    : USINT := 1;
      tock : BOOL  := 0;
  END_VAR
  IF NOT RESET AND tock = NOT TICK THEN
      Data[j]   := IN1;
      Data[j+1] := IN2;
      Data[j+2] := IN3;
      Data[j+3] := IN4;
      Data[j+4] := IN5;
      j := j + 5;
      tock := TICK;
  ELSE
      j := 1;
      tock := 0;
  END_IF;
  Finished := (j > 20);
END_FUNCTION_BLOCK

PROGRAM Boiler
  VAR
    Data  : ARRAY[1..20] OF BOOL;
    Ready : BOOL;
    CollectInput : F_CollectInput;
  END_VAR
  VAR
    TICK     AT %IX1.0 : BOOL;
    IN1      AT %IX0.3 : BOOL;
    IN2      AT %IX0.4 : BOOL;
    IN3      AT %IX0.5 : BOOL;
    IN4      AT %IX0.6 : BOOL;
    IN5      AT %IX0.7 : BOOL;
    OutReady AT %QX0.0 : BOOL := FALSE;
    FeedNext AT %QX0.1 : BOOL := FALSE;
    Out      AT %QX0.2 : BOOL;
  END_VAR
  CollectInput(TICK:=TICK, IN1:=IN1, IN2:=IN2, IN3:=IN3, IN4:=IN4, IN5:=IN5);
  Ready := CollectInput.Finished;
  FeedNext := 1;
  IF Ready THEN
    Out := (((((((((((((((((NOT ((((NOT Data[2]) AND (NOT Data[1])) AND (NOT Data[4])) AND (NOT Data[8]))) OR Data[3]) AND ((NOT (((Data[2] AND (NOT Data[1])) AND (NOT Data[4])) AND (NOT Data[8]))) OR Data[6])) AND ((NOT ((((NOT Data[2]) AND Data[1]) AND (NOT Data[4])) AND (NOT Data[8]))) OR Data[7])) AND ((NOT (((Data[2] AND Data[1]) AND (NOT Data[4])) AND (NOT Data[8]))) OR Data[10])) AND ((NOT ((((NOT Data[2]) AND (NOT Data[1])) AND Data[4]) AND (NOT Data[8]))) OR Data[9])) AND ((NOT (((Data[2] AND (NOT Data[1])) AND Data[4]) AND (NOT Data[8]))) OR Data[5])) AND ((NOT ((((NOT Data[2]) AND Data[1]) AND Data[4]) AND (NOT Data[8]))) OR Data[12])) AND ((NOT (((Data[2] AND Data[1]) AND Data[4]) AND (NOT Data[8]))) OR Data[13])) AND ((NOT ((((NOT Data[2]) AND (NOT Data[1])) AND (NOT Data[4])) AND Data[8])) OR Data[15])) AND ((NOT (((Data[2] AND (NOT Data[1])) AND (NOT Data[4])) AND Data[8])) OR Data[16])) AND ((NOT ((((NOT Data[2]) AND Data[1]) AND (NOT Data[4])) AND Data[8])) OR Data[17])) AND ((NOT (((Data[2] AND Data[1]) AND (NOT Data[4])) AND Data[8])) OR Data[11])) AND ((NOT ((((NOT Data[2]) AND (NOT Data[1])) AND Data[4]) AND Data[8])) OR Data[18])) AND ((NOT (((Data[2] AND (NOT Data[1])) AND Data[4]) AND Data[8])) OR Data[19])) AND ((NOT ((((NOT Data[2]) AND Data[1]) AND Data[4]) AND Data[8])) OR Data[14])) AND ((NOT (((Data[2] AND Data[1]) AND Data[4]) AND Data[8])) OR Data[20]));
    OutReady := 1;
    CollectInput(RESET:=TRUE);
  END_IF;
END_PROGRAM

CONFIGURATION Config0
  RESOURCE Res0 ON PLC
    TASK task0(INTERVAL := T#20ms,PRIORITY := 0);
    PROGRAM instance0 WITH task0 : Boiler;
  END_RESOURCE
END_CONFIGURATION

(* ---- 4-MUX_knelt-salve-hosed.st ---- *)
(*
This code implements a shuffled multiplexer with 4 control bits.
The control bits are: Data[N1], Data[N2], Data[N9], Data[N3]
The input bits are: Data[N4], Data[N5], Data[N6], Data[N7], Data[N8], Data[N11], Data[N14], Data[N10], Data[N12], Data[N13], Data[N15], Data[N17], Data[N19], Data[N16], Data[N20], Data[N18]

The symbolic expression is:
((((((((((((((((!((((!(IN1)) & (!(IN2))) & (!(IN9))) & (!(IN3)))) | IN4) & ((!(((IN1 & (!(IN2))) & (!(IN9))) & (!(IN3)))) | IN5)) & ((!((((!(IN1)) & IN2) & (!(IN9))) & (!(IN3)))) | IN6)) & ((!(((IN1 & IN2) & (!(IN9))) & (!(IN3)))) | IN7)) & ((!((((!(IN1)) & (!(IN2))) & IN9) & (!(IN3)))) | IN8)) & ((!(((IN1 & (!(IN2))) & IN9) & (!(IN3)))) | IN11)) & ((!((((!(IN1)) & IN2) & IN9) & (!(IN3)))) | IN14)) & ((!(((IN1 & IN2) & IN9) & (!(IN3)))) | IN10)) & ((!((((!(IN1)) & (!(IN2))) & (!(IN9))) & IN3)) | IN12)) & ((!(((IN1 & (!(IN2))) & (!(IN9))) & IN3)) | IN13)) & ((!((((!(IN1)) & IN2) & (!(IN9))) & IN3)) | IN15)) & ((!(((IN1 & IN2) & (!(IN9))) & IN3)) | IN17)) & ((!((((!(IN1)) & (!(IN2))) & IN9) & IN3)) | IN19)) & ((!(((IN1 & (!(IN2))) & IN9) & IN3)) | IN16)) & ((!((((!(IN1)) & IN2) & IN9) & IN3)) | IN20)) & ((!(((IN1 & IN2) & IN9) & IN3)) | IN18)

*)

FUNCTION_BLOCK F_CollectInput
  VAR_IN_OUT
      Data : ARRAY[1..20] OF BOOL;
  END_VAR
  VAR_INPUT
      TICK  : BOOL := 0;
      IN1   : BOOL := 0;
      IN2   : BOOL := 0;
      IN3   : BOOL := 0;
      IN4   : BOOL := 0;
      IN5   : BOOL := 0;
      RESET : BOOL := FALSE;
  END_VAR
  VAR_OUTPUT
      Finished : BOOL;
  END_VAR
  VAR
      j    : USINT := 1;
      tock : BOOL  := 0;
  END_VAR
  IF NOT RESET AND tock = NOT TICK THEN
      Data[j]   := IN1;
      Data[j+1] := IN2;
      Data[j+2] := IN3;
      Data[j+3] := IN4;
      Data[j+4] := IN5;
      j := j + 5;
      tock := TICK;
  ELSE
      j := 1;
      tock := 0;
  END_IF;
  Finished := (j > 20);
END_FUNCTION_BLOCK

PROGRAM Boiler
  VAR
    Data  : ARRAY[1..20] OF BOOL;
    Ready : BOOL;
    CollectInput : F_CollectInput;
  END_VAR
  VAR
    TICK     AT %IX1.0 : BOOL;
    IN1      AT %IX0.3 : BOOL;
    IN2      AT %IX0.4 : BOOL;
    IN3      AT %IX0.5 : BOOL;
    IN4      AT %IX0.6 : BOOL;
    IN5      AT %IX0.7 : BOOL;
    OutReady AT %QX0.0 : BOOL := FALSE;
    FeedNext AT %QX0.1 : BOOL := FALSE;
    Out      AT %QX0.2 : BOOL;
  END_VAR
  CollectInput(TICK:=TICK, IN1:=IN1, IN2:=IN2, IN3:=IN3, IN4:=IN4, IN5:=IN5);
  Ready := CollectInput.Finished;
  FeedNext := 1;
  IF Ready THEN
    Out := (((((((((((((((((NOT ((((NOT Data[1]) AND (NOT Data[2])) AND (NOT Data[9])) AND (NOT Data[3]))) OR Data[4]) AND ((NOT (((Data[1] AND (NOT Data[2])) AND (NOT Data[9])) AND (NOT Data[3]))) OR Data[5])) AND ((NOT ((((NOT Data[1]) AND Data[2]) AND (NOT Data[9])) AND (NOT Data[3]))) OR Data[6])) AND ((NOT (((Data[1] AND Data[2]) AND (NOT Data[9])) AND (NOT Data[3]))) OR Data[7])) AND ((NOT ((((NOT Data[1]) AND (NOT Data[2])) AND Data[9]) AND (NOT Data[3]))) OR Data[8])) AND ((NOT (((Data[1] AND (NOT Data[2])) AND Data[9]) AND (NOT Data[3]))) OR Data[11])) AND ((NOT ((((NOT Data[1]) AND Data[2]) AND Data[9]) AND (NOT Data[3]))) OR Data[14])) AND ((NOT (((Data[1] AND Data[2]) AND Data[9]) AND (NOT Data[3]))) OR Data[10])) AND ((NOT ((((NOT Data[1]) AND (NOT Data[2])) AND (NOT Data[9])) AND Data[3])) OR Data[12])) AND ((NOT (((Data[1] AND (NOT Data[2])) AND (NOT Data[9])) AND Data[3])) OR Data[13])) AND ((NOT ((((NOT Data[1]) AND Data[2]) AND (NOT Data[9])) AND Data[3])) OR Data[15])) AND ((NOT (((Data[1] AND Data[2]) AND (NOT Data[9])) AND Data[3])) OR Data[17])) AND ((NOT ((((NOT Data[1]) AND (NOT Data[2])) AND Data[9]) AND Data[3])) OR Data[19])) AND ((NOT (((Data[1] AND (NOT Data[2])) AND Data[9]) AND Data[3])) OR Data[16])) AND ((NOT ((((NOT Data[1]) AND Data[2]) AND Data[9]) AND Data[3])) OR Data[20])) AND ((NOT (((Data[1] AND Data[2]) AND Data[9]) AND Data[3])) OR Data[18]));
    OutReady := 1;
    CollectInput(RESET:=TRUE);
  END_IF;
END_PROGRAM

CONFIGURATION Config0
  RESOURCE Res0 ON PLC
    TASK task0(INTERVAL := T#20ms,PRIORITY := 0);
    PROGRAM instance0 WITH task0 : Boiler;
  END_RESOURCE
END_CONFIGURATION

(* ---- 4-MUX_lames-cruds-cords.st ---- *)
(*
This code implements a shuffled multiplexer with 4 control bits.
The control bits are: Data[N1], Data[N2], Data[N3], Data[N4]
The input bits are: Data[N7], Data[N5], Data[N9], Data[N8], Data[N6], Data[N10], Data[N12], Data[N11], Data[N14], Data[N13], Data[N16], Data[N17], Data[N15], Data[N18], Data[N19], Data[N20]

The symbolic expression is:
((((((((((((((((!((((!(IN1)) & (!(IN2))) & (!(IN3))) & (!(IN4)))) | IN7) & ((!(((IN1 & (!(IN2))) & (!(IN3))) & (!(IN4)))) | IN5)) & ((!((((!(IN1)) & IN2) & (!(IN3))) & (!(IN4)))) | IN9)) & ((!(((IN1 & IN2) & (!(IN3))) & (!(IN4)))) | IN8)) & ((!((((!(IN1)) & (!(IN2))) & IN3) & (!(IN4)))) | IN6)) & ((!(((IN1 & (!(IN2))) & IN3) & (!(IN4)))) | IN10)) & ((!((((!(IN1)) & IN2) & IN3) & (!(IN4)))) | IN12)) & ((!(((IN1 & IN2) & IN3) & (!(IN4)))) | IN11)) & ((!((((!(IN1)) & (!(IN2))) & (!(IN3))) & IN4)) | IN14)) & ((!(((IN1 & (!(IN2))) & (!(IN3))) & IN4)) | IN13)) & ((!((((!(IN1)) & IN2) & (!(IN3))) & IN4)) | IN16)) & ((!(((IN1 & IN2) & (!(IN3))) & IN4)) | IN17)) & ((!((((!(IN1)) & (!(IN2))) & IN3) & IN4)) | IN15)) & ((!(((IN1 & (!(IN2))) & IN3) & IN4)) | IN18)) & ((!((((!(IN1)) & IN2) & IN3) & IN4)) | IN19)) & ((!(((IN1 & IN2) & IN3) & IN4)) | IN20)

*)

FUNCTION_BLOCK F_CollectInput
  VAR_IN_OUT
      Data : ARRAY[1..20] OF BOOL;
  END_VAR
  VAR_INPUT
      TICK  : BOOL := 0;
      IN1   : BOOL := 0;
      IN2   : BOOL := 0;
      IN3   : BOOL := 0;
      IN4   : BOOL := 0;
      IN5   : BOOL := 0;
      RESET : BOOL := FALSE;
  END_VAR
  VAR_OUTPUT
      Finished : BOOL;
  END_VAR
  VAR
      j    : USINT := 1;
      tock : BOOL  := 0;
  END_VAR
  IF NOT RESET AND tock = NOT TICK THEN
      Data[j]   := IN1;
      Data[j+1] := IN2;
      Data[j+2] := IN3;
      Data[j+3] := IN4;
      Data[j+4] := IN5;
      j := j + 5;
      tock := TICK;
  ELSE
      j := 1;
      tock := 0;
  END_IF;
  Finished := (j > 20);
END_FUNCTION_BLOCK

PROGRAM Boiler
  VAR
    Data  : ARRAY[1..20] OF BOOL;
    Ready : BOOL;
    CollectInput : F_CollectInput;
  END_VAR
  VAR
    TICK     AT %IX1.0 : BOOL;
    IN1      AT %IX0.3 : BOOL;
    IN2      AT %IX0.4 : BOOL;
    IN3      AT %IX0.5 : BOOL;
    IN4      AT %IX0.6 : BOOL;
    IN5      AT %IX0.7 : BOOL;
    OutReady AT %QX0.0 : BOOL := FALSE;
    FeedNext AT %QX0.1 : BOOL := FALSE;
    Out      AT %QX0.2 : BOOL;
  END_VAR
  CollectInput(TICK:=TICK, IN1:=IN1, IN2:=IN2, IN3:=IN3, IN4:=IN4, IN5:=IN5);
  Ready := CollectInput.Finished;
  FeedNext := 1;
  IF Ready THEN
    Out := (((((((((((((((((NOT ((((NOT Data[1]) AND (NOT Data[2])) AND (NOT Data[3])) AND (NOT Data[4]))) OR Data[7]) AND ((NOT (((Data[1] AND (NOT Data[2])) AND (NOT Data[3])) AND (NOT Data[4]))) OR Data[5])) AND ((NOT ((((NOT Data[1]) AND Data[2]) AND (NOT Data[3])) AND (NOT Data[4]))) OR Data[9])) AND ((NOT (((Data[1] AND Data[2]) AND (NOT Data[3])) AND (NOT Data[4]))) OR Data[8])) AND ((NOT ((((NOT Data[1]) AND (NOT Data[2])) AND Data[3]) AND (NOT Data[4]))) OR Data[6])) AND ((NOT (((Data[1] AND (NOT Data[2])) AND Data[3]) AND (NOT Data[4]))) OR Data[10])) AND ((NOT ((((NOT Data[1]) AND Data[2]) AND Data[3]) AND (NOT Data[4]))) OR Data[12])) AND ((NOT (((Data[1] AND Data[2]) AND Data[3]) AND (NOT Data[4]))) OR Data[11])) AND ((NOT ((((NOT Data[1]) AND (NOT Data[2])) AND (NOT Data[3])) AND Data[4])) OR Data[14])) AND ((NOT (((Data[1] AND (NOT Data[2])) AND (NOT Data[3])) AND Data[4])) OR Data[13])) AND ((NOT ((((NOT Data[1]) AND Data[2]) AND (NOT Data[3])) AND Data[4])) OR Data[16])) AND ((NOT (((Data[1] AND Data[2]) AND (NOT Data[3])) AND Data[4])) OR Data[17])) AND ((NOT ((((NOT Data[1]) AND (NOT Data[2])) AND Data[3]) AND Data[4])) OR Data[15])) AND ((NOT (((Data[1] AND (NOT Data[2])) AND Data[3]) AND Data[4])) OR Data[18])) AND ((NOT ((((NOT Data[1]) AND Data[2]) AND Data[3]) AND Data[4])) OR Data[19])) AND ((NOT (((Data[1] AND Data[2]) AND Data[3]) AND Data[4])) OR Data[20]));
    OutReady := 1;
    CollectInput(RESET:=TRUE);
  END_IF;
END_PROGRAM

CONFIGURATION Config0
  RESOURCE Res0 ON PLC
    TASK task0(INTERVAL := T#20ms,PRIORITY := 0);
    PROGRAM instance0 WITH task0 : Boiler;
  END_RESOURCE
END_CONFIGURATION

(* ---- 4-MUX_leaps-lived-tweed.st ---- *)
(*
This code implements a shuffled multiplexer with 4 control bits.
The control bits are: Data[N4], Data[N1], Data[N5], Data[N2]
The input bits are: Data[N6], Data[N3], Data[N7], Data[N8], Data[N9], Data[N13], Data[N10], Data[N11], Data[N14], Data[N16], Data[N12], Data[N15], Data[N20], Data[N18], Data[N17], Data[N19]

The symbolic expression is:
((((((((((((((((!((((!(IN4)) & (!(IN1))) & (!(IN5))) & (!(IN2)))) | IN6) & ((!(((IN4 & (!(IN1))) & (!(IN5))) & (!(IN2)))) | IN3)) & ((!((((!(IN4)) & IN1) & (!(IN5))) & (!(IN2)))) | IN7)) & ((!(((IN4 & IN1) & (!(IN5))) & (!(IN2)))) | IN8)) & ((!((((!(IN4)) & (!(IN1))) & IN5) & (!(IN2)))) | IN9)) & ((!(((IN4 & (!(IN1))) & IN5) & (!(IN2)))) | IN13)) & ((!((((!(IN4)) & IN1) & IN5) & (!(IN2)))) | IN10)) & ((!(((IN4 & IN1) & IN5) & (!(IN2)))) | IN11)) & ((!((((!(IN4)) & (!(IN1))) & (!(IN5))) & IN2)) | IN14)) & ((!(((IN4 & (!(IN1))) & (!(IN5))) & IN2)) | IN16)) & ((!((((!(IN4)) & IN1) & (!(IN5))) & IN2)) | IN12)) & ((!(((IN4 & IN1) & (!(IN5))) & IN2)) | IN15)) & ((!((((!(IN4)) & (!(IN1))) & IN5) & IN2)) | IN20)) & ((!(((IN4 & (!(IN1))) & IN5) & IN2)) | IN18)) & ((!((((!(IN4)) & IN1) & IN5) & IN2)) | IN17)) & ((!(((IN4 & IN1) & IN5) & IN2)) | IN19)

*)

FUNCTION_BLOCK F_CollectInput
  VAR_IN_OUT
      Data : ARRAY[1..20] OF BOOL;
  END_VAR
  VAR_INPUT
      TICK  : BOOL := 0;
      IN1   : BOOL := 0;
      IN2   : BOOL := 0;
      IN3   : BOOL := 0;
      IN4   : BOOL := 0;
      IN5   : BOOL := 0;
      RESET : BOOL := FALSE;
  END_VAR
  VAR_OUTPUT
      Finished : BOOL;
  END_VAR
  VAR
      j    : USINT := 1;
      tock : BOOL  := 0;
  END_VAR
  IF NOT RESET AND tock = NOT TICK THEN
      Data[j]   := IN1;
      Data[j+1] := IN2;
      Data[j+2] := IN3;
      Data[j+3] := IN4;
      Data[j+4] := IN5;
      j := j + 5;
      tock := TICK;
  ELSE
      j := 1;
      tock := 0;
  END_IF;
  Finished := (j > 20);
END_FUNCTION_BLOCK

PROGRAM Boiler
  VAR
    Data  : ARRAY[1..20] OF BOOL;
    Ready : BOOL;
    CollectInput : F_CollectInput;
  END_VAR
  VAR
    TICK     AT %IX1.0 : BOOL;
    IN1      AT %IX0.3 : BOOL;
    IN2      AT %IX0.4 : BOOL;
    IN3      AT %IX0.5 : BOOL;
    IN4      AT %IX0.6 : BOOL;
    IN5      AT %IX0.7 : BOOL;
    OutReady AT %QX0.0 : BOOL := FALSE;
    FeedNext AT %QX0.1 : BOOL := FALSE;
    Out      AT %QX0.2 : BOOL;
  END_VAR
  CollectInput(TICK:=TICK, IN1:=IN1, IN2:=IN2, IN3:=IN3, IN4:=IN4, IN5:=IN5);
  Ready := CollectInput.Finished;
  FeedNext := 1;
  IF Ready THEN
    Out := (((((((((((((((((NOT ((((NOT Data[4]) AND (NOT Data[1])) AND (NOT Data[5])) AND (NOT Data[2]))) OR Data[6]) AND ((NOT (((Data[4] AND (NOT Data[1])) AND (NOT Data[5])) AND (NOT Data[2]))) OR Data[3])) AND ((NOT ((((NOT Data[4]) AND Data[1]) AND (NOT Data[5])) AND (NOT Data[2]))) OR Data[7])) AND ((NOT (((Data[4] AND Data[1]) AND (NOT Data[5])) AND (NOT Data[2]))) OR Data[8])) AND ((NOT ((((NOT Data[4]) AND (NOT Data[1])) AND Data[5]) AND (NOT Data[2]))) OR Data[9])) AND ((NOT (((Data[4] AND (NOT Data[1])) AND Data[5]) AND (NOT Data[2]))) OR Data[13])) AND ((NOT ((((NOT Data[4]) AND Data[1]) AND Data[5]) AND (NOT Data[2]))) OR Data[10])) AND ((NOT (((Data[4] AND Data[1]) AND Data[5]) AND (NOT Data[2]))) OR Data[11])) AND ((NOT ((((NOT Data[4]) AND (NOT Data[1])) AND (NOT Data[5])) AND Data[2])) OR Data[14])) AND ((NOT (((Data[4] AND (NOT Data[1])) AND (NOT Data[5])) AND Data[2])) OR Data[16])) AND ((NOT ((((NOT Data[4]) AND Data[1]) AND (NOT Data[5])) AND Data[2])) OR Data[12])) AND ((NOT (((Data[4] AND Data[1]) AND (NOT Data[5])) AND Data[2])) OR Data[15])) AND ((NOT ((((NOT Data[4]) AND (NOT Data[1])) AND Data[5]) AND Data[2])) OR Data[20])) AND ((NOT (((Data[4] AND (NOT Data[1])) AND Data[5]) AND Data[2])) OR Data[18])) AND ((NOT ((((NOT Data[4]) AND Data[1]) AND Data[5]) AND Data[2])) OR Data[17])) AND ((NOT (((Data[4] AND Data[1]) AND Data[5]) AND Data[2])) OR Data[19]));
    OutReady := 1;
    CollectInput(RESET:=TRUE);
  END_IF;
END_PROGRAM

CONFIGURATION Config0
  RESOURCE Res0 ON PLC
    TASK task0(INTERVAL := T#20ms,PRIORITY := 0);
    PROGRAM instance0 WITH task0 : Boiler;
  END_RESOURCE
END_CONFIGURATION

(* ---- 4-MUX_lives-satyr-sappy.st ---- *)
(*
This code implements a shuffled multiplexer with 4 control bits.
The control bits are: Data[N3], Data[N1], Data[N2], Data[N4]
The input bits are: Data[N5], Data[N8], Data[N6], Data[N7], Data[N9], Data[N13], Data[N11], Data[N14], Data[N10], Data[N16], Data[N18], Data[N17], Data[N19], Data[N20], Data[N15], Data[N12]

The symbolic expression is:
((((((((((((((((!((((!(IN3)) & (!(IN1))) & (!(IN2))) & (!(IN4)))) | IN5) & ((!(((IN3 & (!(IN1))) & (!(IN2))) & (!(IN4)))) | IN8)) & ((!((((!(IN3)) & IN1) & (!(IN2))) & (!(IN4)))) | IN6)) & ((!(((IN3 & IN1) & (!(IN2))) & (!(IN4)))) | IN7)) & ((!((((!(IN3)) & (!(IN1))) & IN2) & (!(IN4)))) | IN9)) & ((!(((IN3 & (!(IN1))) & IN2) & (!(IN4)))) | IN13)) & ((!((((!(IN3)) & IN1) & IN2) & (!(IN4)))) | IN11)) & ((!(((IN3 & IN1) & IN2) & (!(IN4)))) | IN14)) & ((!((((!(IN3)) & (!(IN1))) & (!(IN2))) & IN4)) | IN10)) & ((!(((IN3 & (!(IN1))) & (!(IN2))) & IN4)) | IN16)) & ((!((((!(IN3)) & IN1) & (!(IN2))) & IN4)) | IN18)) & ((!(((IN3 & IN1) & (!(IN2))) & IN4)) | IN17)) & ((!((((!(IN3)) & (!(IN1))) & IN2) & IN4)) | IN19)) & ((!(((IN3 & (!(IN1))) & IN2) & IN4)) | IN20)) & ((!((((!(IN3)) & IN1) & IN2) & IN4)) | IN15)) & ((!(((IN3 & IN1) & IN2) & IN4)) | IN12)

*)

FUNCTION_BLOCK F_CollectInput
  VAR_IN_OUT
      Data : ARRAY[1..20] OF BOOL;
  END_VAR
  VAR_INPUT
      TICK  : BOOL := 0;
      IN1   : BOOL := 0;
      IN2   : BOOL := 0;
      IN3   : BOOL := 0;
      IN4   : BOOL := 0;
      IN5   : BOOL := 0;
      RESET : BOOL := FALSE;
  END_VAR
  VAR_OUTPUT
      Finished : BOOL;
  END_VAR
  VAR
      j    : USINT := 1;
      tock : BOOL  := 0;
  END_VAR
  IF NOT RESET AND tock = NOT TICK THEN
      Data[j]   := IN1;
      Data[j+1] := IN2;
      Data[j+2] := IN3;
      Data[j+3] := IN4;
      Data[j+4] := IN5;
      j := j + 5;
      tock := TICK;
  ELSE
      j := 1;
      tock := 0;
  END_IF;
  Finished := (j > 20);
END_FUNCTION_BLOCK

PROGRAM Boiler
  VAR
    Data  : ARRAY[1..20] OF BOOL;
    Ready : BOOL;
    CollectInput : F_CollectInput;
  END_VAR
  VAR
    TICK     AT %IX1.0 : BOOL;
    IN1      AT %IX0.3 : BOOL;
    IN2      AT %IX0.4 : BOOL;
    IN3      AT %IX0.5 : BOOL;
    IN4      AT %IX0.6 : BOOL;
    IN5      AT %IX0.7 : BOOL;
    OutReady AT %QX0.0 : BOOL := FALSE;
    FeedNext AT %QX0.1 : BOOL := FALSE;
    Out      AT %QX0.2 : BOOL;
  END_VAR
  CollectInput(TICK:=TICK, IN1:=IN1, IN2:=IN2, IN3:=IN3, IN4:=IN4, IN5:=IN5);
  Ready := CollectInput.Finished;
  FeedNext := 1;
  IF Ready THEN
    Out := (((((((((((((((((NOT ((((NOT Data[3]) AND (NOT Data[1])) AND (NOT Data[2])) AND (NOT Data[4]))) OR Data[5]) AND ((NOT (((Data[3] AND (NOT Data[1])) AND (NOT Data[2])) AND (NOT Data[4]))) OR Data[8])) AND ((NOT ((((NOT Data[3]) AND Data[1]) AND (NOT Data[2])) AND (NOT Data[4]))) OR Data[6])) AND ((NOT (((Data[3] AND Data[1]) AND (NOT Data[2])) AND (NOT Data[4]))) OR Data[7])) AND ((NOT ((((NOT Data[3]) AND (NOT Data[1])) AND Data[2]) AND (NOT Data[4]))) OR Data[9])) AND ((NOT (((Data[3] AND (NOT Data[1])) AND Data[2]) AND (NOT Data[4]))) OR Data[13])) AND ((NOT ((((NOT Data[3]) AND Data[1]) AND Data[2]) AND (NOT Data[4]))) OR Data[11])) AND ((NOT (((Data[3] AND Data[1]) AND Data[2]) AND (NOT Data[4]))) OR Data[14])) AND ((NOT ((((NOT Data[3]) AND (NOT Data[1])) AND (NOT Data[2])) AND Data[4])) OR Data[10])) AND ((NOT (((Data[3] AND (NOT Data[1])) AND (NOT Data[2])) AND Data[4])) OR Data[16])) AND ((NOT ((((NOT Data[3]) AND Data[1]) AND (NOT Data[2])) AND Data[4])) OR Data[18])) AND ((NOT (((Data[3] AND Data[1]) AND (NOT Data[2])) AND Data[4])) OR Data[17])) AND ((NOT ((((NOT Data[3]) AND (NOT Data[1])) AND Data[2]) AND Data[4])) OR Data[19])) AND ((NOT (((Data[3] AND (NOT Data[1])) AND Data[2]) AND Data[4])) OR Data[20])) AND ((NOT ((((NOT Data[3]) AND Data[1]) AND Data[2]) AND Data[4])) OR Data[15])) AND ((NOT (((Data[3] AND Data[1]) AND Data[2]) AND Data[4])) OR Data[12]));
    OutReady := 1;
    CollectInput(RESET:=TRUE);
  END_IF;
END_PROGRAM

CONFIGURATION Config0
  RESOURCE Res0 ON PLC
    TASK task0(INTERVAL := T#20ms,PRIORITY := 0);
    PROGRAM instance0 WITH task0 : Boiler;
  END_RESOURCE
END_CONFIGURATION

(* ---- 4-MUX_loppy-hasps-slung.st ---- *)
(*
This code implements a shuffled multiplexer with 4 control bits.
The control bits are: Data[N3], Data[N1], Data[N6], Data[N8]
The input bits are: Data[N4], Data[N2], Data[N7], Data[N9], Data[N5], Data[N13], Data[N10], Data[N11], Data[N12], Data[N14], Data[N15], Data[N16], Data[N17], Data[N18], Data[N20], Data[N19]

The symbolic expression is:
((((((((((((((((!((((!(IN3)) & (!(IN1))) & (!(IN6))) & (!(IN8)))) | IN4) & ((!(((IN3 & (!(IN1))) & (!(IN6))) & (!(IN8)))) | IN2)) & ((!((((!(IN3)) & IN1) & (!(IN6))) & (!(IN8)))) | IN7)) & ((!(((IN3 & IN1) & (!(IN6))) & (!(IN8)))) | IN9)) & ((!((((!(IN3)) & (!(IN1))) & IN6) & (!(IN8)))) | IN5)) & ((!(((IN3 & (!(IN1))) & IN6) & (!(IN8)))) | IN13)) & ((!((((!(IN3)) & IN1) & IN6) & (!(IN8)))) | IN10)) & ((!(((IN3 & IN1) & IN6) & (!(IN8)))) | IN11)) & ((!((((!(IN3)) & (!(IN1))) & (!(IN6))) & IN8)) | IN12)) & ((!(((IN3 & (!(IN1))) & (!(IN6))) & IN8)) | IN14)) & ((!((((!(IN3)) & IN1) & (!(IN6))) & IN8)) | IN15)) & ((!(((IN3 & IN1) & (!(IN6))) & IN8)) | IN16)) & ((!((((!(IN3)) & (!(IN1))) & IN6) & IN8)) | IN17)) & ((!(((IN3 & (!(IN1))) & IN6) & IN8)) | IN18)) & ((!((((!(IN3)) & IN1) & IN6) & IN8)) | IN20)) & ((!(((IN3 & IN1) & IN6) & IN8)) | IN19)

*)

FUNCTION_BLOCK F_CollectInput
  VAR_IN_OUT
      Data : ARRAY[1..20] OF BOOL;
  END_VAR
  VAR_INPUT
      TICK  : BOOL := 0;
      IN1   : BOOL := 0;
      IN2   : BOOL := 0;
      IN3   : BOOL := 0;
      IN4   : BOOL := 0;
      IN5   : BOOL := 0;
      RESET : BOOL := FALSE;
  END_VAR
  VAR_OUTPUT
      Finished : BOOL;
  END_VAR
  VAR
      j    : USINT := 1;
      tock : BOOL  := 0;
  END_VAR
  IF NOT RESET AND tock = NOT TICK THEN
      Data[j]   := IN1;
      Data[j+1] := IN2;
      Data[j+2] := IN3;
      Data[j+3] := IN4;
      Data[j+4] := IN5;
      j := j + 5;
      tock := TICK;
  ELSE
      j := 1;
      tock := 0;
  END_IF;
  Finished := (j > 20);
END_FUNCTION_BLOCK

PROGRAM Boiler
  VAR
    Data  : ARRAY[1..20] OF BOOL;
    Ready : BOOL;
    CollectInput : F_CollectInput;
  END_VAR
  VAR
    TICK     AT %IX1.0 : BOOL;
    IN1      AT %IX0.3 : BOOL;
    IN2      AT %IX0.4 : BOOL;
    IN3      AT %IX0.5 : BOOL;
    IN4      AT %IX0.6 : BOOL;
    IN5      AT %IX0.7 : BOOL;
    OutReady AT %QX0.0 : BOOL := FALSE;
    FeedNext AT %QX0.1 : BOOL := FALSE;
    Out      AT %QX0.2 : BOOL;
  END_VAR
  CollectInput(TICK:=TICK, IN1:=IN1, IN2:=IN2, IN3:=IN3, IN4:=IN4, IN5:=IN5);
  Ready := CollectInput.Finished;
  FeedNext := 1;
  IF Ready THEN
    Out := (((((((((((((((((NOT ((((NOT Data[3]) AND (NOT Data[1])) AND (NOT Data[6])) AND (NOT Data[8]))) OR Data[4]) AND ((NOT (((Data[3] AND (NOT Data[1])) AND (NOT Data[6])) AND (NOT Data[8]))) OR Data[2])) AND ((NOT ((((NOT Data[3]) AND Data[1]) AND (NOT Data[6])) AND (NOT Data[8]))) OR Data[7])) AND ((NOT (((Data[3] AND Data[1]) AND (NOT Data[6])) AND (NOT Data[8]))) OR Data[9])) AND ((NOT ((((NOT Data[3]) AND (NOT Data[1])) AND Data[6]) AND (NOT Data[8]))) OR Data[5])) AND ((NOT (((Data[3] AND (NOT Data[1])) AND Data[6]) AND (NOT Data[8]))) OR Data[13])) AND ((NOT ((((NOT Data[3]) AND Data[1]) AND Data[6]) AND (NOT Data[8]))) OR Data[10])) AND ((NOT (((Data[3] AND Data[1]) AND Data[6]) AND (NOT Data[8]))) OR Data[11])) AND ((NOT ((((NOT Data[3]) AND (NOT Data[1])) AND (NOT Data[6])) AND Data[8])) OR Data[12])) AND ((NOT (((Data[3] AND (NOT Data[1])) AND (NOT Data[6])) AND Data[8])) OR Data[14])) AND ((NOT ((((NOT Data[3]) AND Data[1]) AND (NOT Data[6])) AND Data[8])) OR Data[15])) AND ((NOT (((Data[3] AND Data[1]) AND (NOT Data[6])) AND Data[8])) OR Data[16])) AND ((NOT ((((NOT Data[3]) AND (NOT Data[1])) AND Data[6]) AND Data[8])) OR Data[17])) AND ((NOT (((Data[3] AND (NOT Data[1])) AND Data[6]) AND Data[8])) OR Data[18])) AND ((NOT ((((NOT Data[3]) AND Data[1]) AND Data[6]) AND Data[8])) OR Data[20])) AND ((NOT (((Data[3] AND Data[1]) AND Data[6]) AND Data[8])) OR Data[19]));
    OutReady := 1;
    CollectInput(RESET:=TRUE);
  END_IF;
END_PROGRAM

CONFIGURATION Config0
  RESOURCE Res0 ON PLC
    TASK task0(INTERVAL := T#20ms,PRIORITY := 0);
    PROGRAM instance0 WITH task0 : Boiler;
  END_RESOURCE
END_CONFIGURATION

(* ---- 4-MUX_lured-dorks-veils.st ---- *)
(*
This code implements a shuffled multiplexer with 4 control bits.
The control bits are: Data[N1], Data[N4], Data[N3], Data[N6]
The input bits are: Data[N2], Data[N7], Data[N5], Data[N8], Data[N12], Data[N10], Data[N13], Data[N9], Data[N15], Data[N11], Data[N14], Data[N17], Data[N16], Data[N20], Data[N19], Data[N18]

The symbolic expression is:
((((((((((((((((!((((!(IN1)) & (!(IN4))) & (!(IN3))) & (!(IN6)))) | IN2) & ((!(((IN1 & (!(IN4))) & (!(IN3))) & (!(IN6)))) | IN7)) & ((!((((!(IN1)) & IN4) & (!(IN3))) & (!(IN6)))) | IN5)) & ((!(((IN1 & IN4) & (!(IN3))) & (!(IN6)))) | IN8)) & ((!((((!(IN1)) & (!(IN4))) & IN3) & (!(IN6)))) | IN12)) & ((!(((IN1 & (!(IN4))) & IN3) & (!(IN6)))) | IN10)) & ((!((((!(IN1)) & IN4) & IN3) & (!(IN6)))) | IN13)) & ((!(((IN1 & IN4) & IN3) & (!(IN6)))) | IN9)) & ((!((((!(IN1)) & (!(IN4))) & (!(IN3))) & IN6)) | IN15)) & ((!(((IN1 & (!(IN4))) & (!(IN3))) & IN6)) | IN11)) & ((!((((!(IN1)) & IN4) & (!(IN3))) & IN6)) | IN14)) & ((!(((IN1 & IN4) & (!(IN3))) & IN6)) | IN17)) & ((!((((!(IN1)) & (!(IN4))) & IN3) & IN6)) | IN16)) & ((!(((IN1 & (!(IN4))) & IN3) & IN6)) | IN20)) & ((!((((!(IN1)) & IN4) & IN3) & IN6)) | IN19)) & ((!(((IN1 & IN4) & IN3) & IN6)) | IN18)

*)

FUNCTION_BLOCK F_CollectInput
  VAR_IN_OUT
      Data : ARRAY[1..20] OF BOOL;
  END_VAR
  VAR_INPUT
      TICK  : BOOL := 0;
      IN1   : BOOL := 0;
      IN2   : BOOL := 0;
      IN3   : BOOL := 0;
      IN4   : BOOL := 0;
      IN5   : BOOL := 0;
      RESET : BOOL := FALSE;
  END_VAR
  VAR_OUTPUT
      Finished : BOOL;
  END_VAR
  VAR
      j    : USINT := 1;
      tock : BOOL  := 0;
  END_VAR
  IF NOT RESET AND tock = NOT TICK THEN
      Data[j]   := IN1;
      Data[j+1] := IN2;
      Data[j+2] := IN3;
      Data[j+3] := IN4;
      Data[j+4] := IN5;
      j := j + 5;
      tock := TICK;
  ELSE
      j := 1;
      tock := 0;
  END_IF;
  Finished := (j > 20);
END_FUNCTION_BLOCK

PROGRAM Boiler
  VAR
    Data  : ARRAY[1..20] OF BOOL;
    Ready : BOOL;
    CollectInput : F_CollectInput;
  END_VAR
  VAR
    TICK     AT %IX1.0 : BOOL;
    IN1      AT %IX0.3 : BOOL;
    IN2      AT %IX0.4 : BOOL;
    IN3      AT %IX0.5 : BOOL;
    IN4      AT %IX0.6 : BOOL;
    IN5      AT %IX0.7 : BOOL;
    OutReady AT %QX0.0 : BOOL := FALSE;
    FeedNext AT %QX0.1 : BOOL := FALSE;
    Out      AT %QX0.2 : BOOL;
  END_VAR
  CollectInput(TICK:=TICK, IN1:=IN1, IN2:=IN2, IN3:=IN3, IN4:=IN4, IN5:=IN5);
  Ready := CollectInput.Finished;
  FeedNext := 1;
  IF Ready THEN
    Out := (((((((((((((((((NOT ((((NOT Data[1]) AND (NOT Data[4])) AND (NOT Data[3])) AND (NOT Data[6]))) OR Data[2]) AND ((NOT (((Data[1] AND (NOT Data[4])) AND (NOT Data[3])) AND (NOT Data[6]))) OR Data[7])) AND ((NOT ((((NOT Data[1]) AND Data[4]) AND (NOT Data[3])) AND (NOT Data[6]))) OR Data[5])) AND ((NOT (((Data[1] AND Data[4]) AND (NOT Data[3])) AND (NOT Data[6]))) OR Data[8])) AND ((NOT ((((NOT Data[1]) AND (NOT Data[4])) AND Data[3]) AND (NOT Data[6]))) OR Data[12])) AND ((NOT (((Data[1] AND (NOT Data[4])) AND Data[3]) AND (NOT Data[6]))) OR Data[10])) AND ((NOT ((((NOT Data[1]) AND Data[4]) AND Data[3]) AND (NOT Data[6]))) OR Data[13])) AND ((NOT (((Data[1] AND Data[4]) AND Data[3]) AND (NOT Data[6]))) OR Data[9])) AND ((NOT ((((NOT Data[1]) AND (NOT Data[4])) AND (NOT Data[3])) AND Data[6])) OR Data[15])) AND ((NOT (((Data[1] AND (NOT Data[4])) AND (NOT Data[3])) AND Data[6])) OR Data[11])) AND ((NOT ((((NOT Data[1]) AND Data[4]) AND (NOT Data[3])) AND Data[6])) OR Data[14])) AND ((NOT (((Data[1] AND Data[4]) AND (NOT Data[3])) AND Data[6])) OR Data[17])) AND ((NOT ((((NOT Data[1]) AND (NOT Data[4])) AND Data[3]) AND Data[6])) OR Data[16])) AND ((NOT (((Data[1] AND (NOT Data[4])) AND Data[3]) AND Data[6])) OR Data[20])) AND ((NOT ((((NOT Data[1]) AND Data[4]) AND Data[3]) AND Data[6])) OR Data[19])) AND ((NOT (((Data[1] AND Data[4]) AND Data[3]) AND Data[6])) OR Data[18]));
    OutReady := 1;
    CollectInput(RESET:=TRUE);
  END_IF;
END_PROGRAM

CONFIGURATION Config0
  RESOURCE Res0 ON PLC
    TASK task0(INTERVAL := T#20ms,PRIORITY := 0);
    PROGRAM instance0 WITH task0 : Boiler;
  END_RESOURCE
END_CONFIGURATION

(* ---- 4-MUX_match-bangs-wises.st ---- *)
(*
This code implements a shuffled multiplexer with 4 control bits.
The control bits are: Data[N7], Data[N3], Data[N11], Data[N4]
The input bits are: Data[N1], Data[N6], Data[N5], Data[N9], Data[N8], Data[N2], Data[N12], Data[N10], Data[N13], Data[N14], Data[N15], Data[N16], Data[N17], Data[N18], Data[N19], Data[N20]

The symbolic expression is:
((((((((((((((((!((((!(IN7)) & (!(IN3))) & (!(IN11))) & (!(IN4)))) | IN1) & ((!(((IN7 & (!(IN3))) & (!(IN11))) & (!(IN4)))) | IN6)) & ((!((((!(IN7)) & IN3) & (!(IN11))) & (!(IN4)))) | IN5)) & ((!(((IN7 & IN3) & (!(IN11))) & (!(IN4)))) | IN9)) & ((!((((!(IN7)) & (!(IN3))) & IN11) & (!(IN4)))) | IN8)) & ((!(((IN7 & (!(IN3))) & IN11) & (!(IN4)))) | IN2)) & ((!((((!(IN7)) & IN3) & IN11) & (!(IN4)))) | IN12)) & ((!(((IN7 & IN3) & IN11) & (!(IN4)))) | IN10)) & ((!((((!(IN7)) & (!(IN3))) & (!(IN11))) & IN4)) | IN13)) & ((!(((IN7 & (!(IN3))) & (!(IN11))) & IN4)) | IN14)) & ((!((((!(IN7)) & IN3) & (!(IN11))) & IN4)) | IN15)) & ((!(((IN7 & IN3) & (!(IN11))) & IN4)) | IN16)) & ((!((((!(IN7)) & (!(IN3))) & IN11) & IN4)) | IN17)) & ((!(((IN7 & (!(IN3))) & IN11) & IN4)) | IN18)) & ((!((((!(IN7)) & IN3) & IN11) & IN4)) | IN19)) & ((!(((IN7 & IN3) & IN11) & IN4)) | IN20)

*)

FUNCTION_BLOCK F_CollectInput
  VAR_IN_OUT
      Data : ARRAY[1..20] OF BOOL;
  END_VAR
  VAR_INPUT
      TICK  : BOOL := 0;
      IN1   : BOOL := 0;
      IN2   : BOOL := 0;
      IN3   : BOOL := 0;
      IN4   : BOOL := 0;
      IN5   : BOOL := 0;
      RESET : BOOL := FALSE;
  END_VAR
  VAR_OUTPUT
      Finished : BOOL;
  END_VAR
  VAR
      j    : USINT := 1;
      tock : BOOL  := 0;
  END_VAR
  IF NOT RESET AND tock = NOT TICK THEN
      Data[j]   := IN1;
      Data[j+1] := IN2;
      Data[j+2] := IN3;
      Data[j+3] := IN4;
      Data[j+4] := IN5;
      j := j + 5;
      tock := TICK;
  ELSE
      j := 1;
      tock := 0;
  END_IF;
  Finished := (j > 20);
END_FUNCTION_BLOCK

PROGRAM Boiler
  VAR
    Data  : ARRAY[1..20] OF BOOL;
    Ready : BOOL;
    CollectInput : F_CollectInput;
  END_VAR
  VAR
    TICK     AT %IX1.0 : BOOL;
    IN1      AT %IX0.3 : BOOL;
    IN2      AT %IX0.4 : BOOL;
    IN3      AT %IX0.5 : BOOL;
    IN4      AT %IX0.6 : BOOL;
    IN5      AT %IX0.7 : BOOL;
    OutReady AT %QX0.0 : BOOL := FALSE;
    FeedNext AT %QX0.1 : BOOL := FALSE;
    Out      AT %QX0.2 : BOOL;
  END_VAR
  CollectInput(TICK:=TICK, IN1:=IN1, IN2:=IN2, IN3:=IN3, IN4:=IN4, IN5:=IN5);
  Ready := CollectInput.Finished;
  FeedNext := 1;
  IF Ready THEN
    Out := (((((((((((((((((NOT ((((NOT Data[7]) AND (NOT Data[3])) AND (NOT Data[11])) AND (NOT Data[4]))) OR Data[1]) AND ((NOT (((Data[7] AND (NOT Data[3])) AND (NOT Data[11])) AND (NOT Data[4]))) OR Data[6])) AND ((NOT ((((NOT Data[7]) AND Data[3]) AND (NOT Data[11])) AND (NOT Data[4]))) OR Data[5])) AND ((NOT (((Data[7] AND Data[3]) AND (NOT Data[11])) AND (NOT Data[4]))) OR Data[9])) AND ((NOT ((((NOT Data[7]) AND (NOT Data[3])) AND Data[11]) AND (NOT Data[4]))) OR Data[8])) AND ((NOT (((Data[7] AND (NOT Data[3])) AND Data[11]) AND (NOT Data[4]))) OR Data[2])) AND ((NOT ((((NOT Data[7]) AND Data[3]) AND Data[11]) AND (NOT Data[4]))) OR Data[12])) AND ((NOT (((Data[7] AND Data[3]) AND Data[11]) AND (NOT Data[4]))) OR Data[10])) AND ((NOT ((((NOT Data[7]) AND (NOT Data[3])) AND (NOT Data[11])) AND Data[4])) OR Data[13])) AND ((NOT (((Data[7] AND (NOT Data[3])) AND (NOT Data[11])) AND Data[4])) OR Data[14])) AND ((NOT ((((NOT Data[7]) AND Data[3]) AND (NOT Data[11])) AND Data[4])) OR Data[15])) AND ((NOT (((Data[7] AND Data[3]) AND (NOT Data[11])) AND Data[4])) OR Data[16])) AND ((NOT ((((NOT Data[7]) AND (NOT Data[3])) AND Data[11]) AND Data[4])) OR Data[17])) AND ((NOT (((Data[7] AND (NOT Data[3])) AND Data[11]) AND Data[4])) OR Data[18])) AND ((NOT ((((NOT Data[7]) AND Data[3]) AND Data[11]) AND Data[4])) OR Data[19])) AND ((NOT (((Data[7] AND Data[3]) AND Data[11]) AND Data[4])) OR Data[20]));
    OutReady := 1;
    CollectInput(RESET:=TRUE);
  END_IF;
END_PROGRAM

CONFIGURATION Config0
  RESOURCE Res0 ON PLC
    TASK task0(INTERVAL := T#20ms,PRIORITY := 0);
    PROGRAM instance0 WITH task0 : Boiler;
  END_RESOURCE
END_CONFIGURATION

(* ---- 4-MUX_meows-scoop-swift.st ---- *)
(*
This code implements a shuffled multiplexer with 4 control bits.
The control bits are: Data[N4], Data[N3], Data[N2], Data[N5]
The input bits are: Data[N1], Data[N7], Data[N12], Data[N6], Data[N8], Data[N9], Data[N13], Data[N15], Data[N10], Data[N11], Data[N14], Data[N17], Data[N18], Data[N20], Data[N16], Data[N19]

The symbolic expression is:
((((((((((((((((!((((!(IN4)) & (!(IN3))) & (!(IN2))) & (!(IN5)))) | IN1) & ((!(((IN4 & (!(IN3))) & (!(IN2))) & (!(IN5)))) | IN7)) & ((!((((!(IN4)) & IN3) & (!(IN2))) & (!(IN5)))) | IN12)) & ((!(((IN4 & IN3) & (!(IN2))) & (!(IN5)))) | IN6)) & ((!((((!(IN4)) & (!(IN3))) & IN2) & (!(IN5)))) | IN8)) & ((!(((IN4 & (!(IN3))) & IN2) & (!(IN5)))) | IN9)) & ((!((((!(IN4)) & IN3) & IN2) & (!(IN5)))) | IN13)) & ((!(((IN4 & IN3) & IN2) & (!(IN5)))) | IN15)) & ((!((((!(IN4)) & (!(IN3))) & (!(IN2))) & IN5)) | IN10)) & ((!(((IN4 & (!(IN3))) & (!(IN2))) & IN5)) | IN11)) & ((!((((!(IN4)) & IN3) & (!(IN2))) & IN5)) | IN14)) & ((!(((IN4 & IN3) & (!(IN2))) & IN5)) | IN17)) & ((!((((!(IN4)) & (!(IN3))) & IN2) & IN5)) | IN18)) & ((!(((IN4 & (!(IN3))) & IN2) & IN5)) | IN20)) & ((!((((!(IN4)) & IN3) & IN2) & IN5)) | IN16)) & ((!(((IN4 & IN3) & IN2) & IN5)) | IN19)

*)

FUNCTION_BLOCK F_CollectInput
  VAR_IN_OUT
      Data : ARRAY[1..20] OF BOOL;
  END_VAR
  VAR_INPUT
      TICK  : BOOL := 0;
      IN1   : BOOL := 0;
      IN2   : BOOL := 0;
      IN3   : BOOL := 0;
      IN4   : BOOL := 0;
      IN5   : BOOL := 0;
      RESET : BOOL := FALSE;
  END_VAR
  VAR_OUTPUT
      Finished : BOOL;
  END_VAR
  VAR
      j    : USINT := 1;
      tock : BOOL  := 0;
  END_VAR
  IF NOT RESET AND tock = NOT TICK THEN
      Data[j]   := IN1;
      Data[j+1] := IN2;
      Data[j+2] := IN3;
      Data[j+3] := IN4;
      Data[j+4] := IN5;
      j := j + 5;
      tock := TICK;
  ELSE
      j := 1;
      tock := 0;
  END_IF;
  Finished := (j > 20);
END_FUNCTION_BLOCK

PROGRAM Boiler
  VAR
    Data  : ARRAY[1..20] OF BOOL;
    Ready : BOOL;
    CollectInput : F_CollectInput;
  END_VAR
  VAR
    TICK     AT %IX1.0 : BOOL;
    IN1      AT %IX0.3 : BOOL;
    IN2      AT %IX0.4 : BOOL;
    IN3      AT %IX0.5 : BOOL;
    IN4      AT %IX0.6 : BOOL;
    IN5      AT %IX0.7 : BOOL;
    OutReady AT %QX0.0 : BOOL := FALSE;
    FeedNext AT %QX0.1 : BOOL := FALSE;
    Out      AT %QX0.2 : BOOL;
  END_VAR
  CollectInput(TICK:=TICK, IN1:=IN1, IN2:=IN2, IN3:=IN3, IN4:=IN4, IN5:=IN5);
  Ready := CollectInput.Finished;
  FeedNext := 1;
  IF Ready THEN
    Out := (((((((((((((((((NOT ((((NOT Data[4]) AND (NOT Data[3])) AND (NOT Data[2])) AND (NOT Data[5]))) OR Data[1]) AND ((NOT (((Data[4] AND (NOT Data[3])) AND (NOT Data[2])) AND (NOT Data[5]))) OR Data[7])) AND ((NOT ((((NOT Data[4]) AND Data[3]) AND (NOT Data[2])) AND (NOT Data[5]))) OR Data[12])) AND ((NOT (((Data[4] AND Data[3]) AND (NOT Data[2])) AND (NOT Data[5]))) OR Data[6])) AND ((NOT ((((NOT Data[4]) AND (NOT Data[3])) AND Data[2]) AND (NOT Data[5]))) OR Data[8])) AND ((NOT (((Data[4] AND (NOT Data[3])) AND Data[2]) AND (NOT Data[5]))) OR Data[9])) AND ((NOT ((((NOT Data[4]) AND Data[3]) AND Data[2]) AND (NOT Data[5]))) OR Data[13])) AND ((NOT (((Data[4] AND Data[3]) AND Data[2]) AND (NOT Data[5]))) OR Data[15])) AND ((NOT ((((NOT Data[4]) AND (NOT Data[3])) AND (NOT Data[2])) AND Data[5])) OR Data[10])) AND ((NOT (((Data[4] AND (NOT Data[3])) AND (NOT Data[2])) AND Data[5])) OR Data[11])) AND ((NOT ((((NOT Data[4]) AND Data[3]) AND (NOT Data[2])) AND Data[5])) OR Data[14])) AND ((NOT (((Data[4] AND Data[3]) AND (NOT Data[2])) AND Data[5])) OR Data[17])) AND ((NOT ((((NOT Data[4]) AND (NOT Data[3])) AND Data[2]) AND Data[5])) OR Data[18])) AND ((NOT (((Data[4] AND (NOT Data[3])) AND Data[2]) AND Data[5])) OR Data[20])) AND ((NOT ((((NOT Data[4]) AND Data[3]) AND Data[2]) AND Data[5])) OR Data[16])) AND ((NOT (((Data[4] AND Data[3]) AND Data[2]) AND Data[5])) OR Data[19]));
    OutReady := 1;
    CollectInput(RESET:=TRUE);
  END_IF;
END_PROGRAM

CONFIGURATION Config0
  RESOURCE Res0 ON PLC
    TASK task0(INTERVAL := T#20ms,PRIORITY := 0);
    PROGRAM instance0 WITH task0 : Boiler;
  END_RESOURCE
END_CONFIGURATION

(* ---- 4-MUX_miked-kinky-hangs.st ---- *)
(*
This code implements a shuffled multiplexer with 4 control bits.
The control bits are: Data[N1], Data[N2], Data[N3], Data[N4]
The input bits are: Data[N7], Data[N6], Data[N5], Data[N8], Data[N9], Data[N11], Data[N12], Data[N13], Data[N16], Data[N10], Data[N15], Data[N14], Data[N18], Data[N17], Data[N19], Data[N20]

The symbolic expression is:
((((((((((((((((!((((!(IN1)) & (!(IN2))) & (!(IN3))) & (!(IN4)))) | IN7) & ((!(((IN1 & (!(IN2))) & (!(IN3))) & (!(IN4)))) | IN6)) & ((!((((!(IN1)) & IN2) & (!(IN3))) & (!(IN4)))) | IN5)) & ((!(((IN1 & IN2) & (!(IN3))) & (!(IN4)))) | IN8)) & ((!((((!(IN1)) & (!(IN2))) & IN3) & (!(IN4)))) | IN9)) & ((!(((IN1 & (!(IN2))) & IN3) & (!(IN4)))) | IN11)) & ((!((((!(IN1)) & IN2) & IN3) & (!(IN4)))) | IN12)) & ((!(((IN1 & IN2) & IN3) & (!(IN4)))) | IN13)) & ((!((((!(IN1)) & (!(IN2))) & (!(IN3))) & IN4)) | IN16)) & ((!(((IN1 & (!(IN2))) & (!(IN3))) & IN4)) | IN10)) & ((!((((!(IN1)) & IN2) & (!(IN3))) & IN4)) | IN15)) & ((!(((IN1 & IN2) & (!(IN3))) & IN4)) | IN14)) & ((!((((!(IN1)) & (!(IN2))) & IN3) & IN4)) | IN18)) & ((!(((IN1 & (!(IN2))) & IN3) & IN4)) | IN17)) & ((!((((!(IN1)) & IN2) & IN3) & IN4)) | IN19)) & ((!(((IN1 & IN2) & IN3) & IN4)) | IN20)

*)

FUNCTION_BLOCK F_CollectInput
  VAR_IN_OUT
      Data : ARRAY[1..20] OF BOOL;
  END_VAR
  VAR_INPUT
      TICK  : BOOL := 0;
      IN1   : BOOL := 0;
      IN2   : BOOL := 0;
      IN3   : BOOL := 0;
      IN4   : BOOL := 0;
      IN5   : BOOL := 0;
      RESET : BOOL := FALSE;
  END_VAR
  VAR_OUTPUT
      Finished : BOOL;
  END_VAR
  VAR
      j    : USINT := 1;
      tock : BOOL  := 0;
  END_VAR
  IF NOT RESET AND tock = NOT TICK THEN
      Data[j]   := IN1;
      Data[j+1] := IN2;
      Data[j+2] := IN3;
      Data[j+3] := IN4;
      Data[j+4] := IN5;
      j := j + 5;
      tock := TICK;
  ELSE
      j := 1;
      tock := 0;
  END_IF;
  Finished := (j > 20);
END_FUNCTION_BLOCK

PROGRAM Boiler
  VAR
    Data  : ARRAY[1..20] OF BOOL;
    Ready : BOOL;
    CollectInput : F_CollectInput;
  END_VAR
  VAR
    TICK     AT %IX1.0 : BOOL;
    IN1      AT %IX0.3 : BOOL;
    IN2      AT %IX0.4 : BOOL;
    IN3      AT %IX0.5 : BOOL;
    IN4      AT %IX0.6 : BOOL;
    IN5      AT %IX0.7 : BOOL;
    OutReady AT %QX0.0 : BOOL := FALSE;
    FeedNext AT %QX0.1 : BOOL := FALSE;
    Out      AT %QX0.2 : BOOL;
  END_VAR
  CollectInput(TICK:=TICK, IN1:=IN1, IN2:=IN2, IN3:=IN3, IN4:=IN4, IN5:=IN5);
  Ready := CollectInput.Finished;
  FeedNext := 1;
  IF Ready THEN
    Out := (((((((((((((((((NOT ((((NOT Data[1]) AND (NOT Data[2])) AND (NOT Data[3])) AND (NOT Data[4]))) OR Data[7]) AND ((NOT (((Data[1] AND (NOT Data[2])) AND (NOT Data[3])) AND (NOT Data[4]))) OR Data[6])) AND ((NOT ((((NOT Data[1]) AND Data[2]) AND (NOT Data[3])) AND (NOT Data[4]))) OR Data[5])) AND ((NOT (((Data[1] AND Data[2]) AND (NOT Data[3])) AND (NOT Data[4]))) OR Data[8])) AND ((NOT ((((NOT Data[1]) AND (NOT Data[2])) AND Data[3]) AND (NOT Data[4]))) OR Data[9])) AND ((NOT (((Data[1] AND (NOT Data[2])) AND Data[3]) AND (NOT Data[4]))) OR Data[11])) AND ((NOT ((((NOT Data[1]) AND Data[2]) AND Data[3]) AND (NOT Data[4]))) OR Data[12])) AND ((NOT (((Data[1] AND Data[2]) AND Data[3]) AND (NOT Data[4]))) OR Data[13])) AND ((NOT ((((NOT Data[1]) AND (NOT Data[2])) AND (NOT Data[3])) AND Data[4])) OR Data[16])) AND ((NOT (((Data[1] AND (NOT Data[2])) AND (NOT Data[3])) AND Data[4])) OR Data[10])) AND ((NOT ((((NOT Data[1]) AND Data[2]) AND (NOT Data[3])) AND Data[4])) OR Data[15])) AND ((NOT (((Data[1] AND Data[2]) AND (NOT Data[3])) AND Data[4])) OR Data[14])) AND ((NOT ((((NOT Data[1]) AND (NOT Data[2])) AND Data[3]) AND Data[4])) OR Data[18])) AND ((NOT (((Data[1] AND (NOT Data[2])) AND Data[3]) AND Data[4])) OR Data[17])) AND ((NOT ((((NOT Data[1]) AND Data[2]) AND Data[3]) AND Data[4])) OR Data[19])) AND ((NOT (((Data[1] AND Data[2]) AND Data[3]) AND Data[4])) OR Data[20]));
    OutReady := 1;
    CollectInput(RESET:=TRUE);
  END_IF;
END_PROGRAM

CONFIGURATION Config0
  RESOURCE Res0 ON PLC
    TASK task0(INTERVAL := T#20ms,PRIORITY := 0);
    PROGRAM instance0 WITH task0 : Boiler;
  END_RESOURCE
END_CONFIGURATION

(* ---- 4-MUX_mucus-otter-clang.st ---- *)
(*
This code implements a shuffled multiplexer with 4 control bits.
The control bits are: Data[N1], Data[N4], Data[N3], Data[N2]
The input bits are: Data[N8], Data[N5], Data[N6], Data[N9], Data[N7], Data[N10], Data[N12], Data[N11], Data[N13], Data[N14], Data[N15], Data[N16], Data[N17], Data[N18], Data[N19], Data[N20]

The symbolic expression is:
((((((((((((((((!((((!(IN1)) & (!(IN4))) & (!(IN3))) & (!(IN2)))) | IN8) & ((!(((IN1 & (!(IN4))) & (!(IN3))) & (!(IN2)))) | IN5)) & ((!((((!(IN1)) & IN4) & (!(IN3))) & (!(IN2)))) | IN6)) & ((!(((IN1 & IN4) & (!(IN3))) & (!(IN2)))) | IN9)) & ((!((((!(IN1)) & (!(IN4))) & IN3) & (!(IN2)))) | IN7)) & ((!(((IN1 & (!(IN4))) & IN3) & (!(IN2)))) | IN10)) & ((!((((!(IN1)) & IN4) & IN3) & (!(IN2)))) | IN12)) & ((!(((IN1 & IN4) & IN3) & (!(IN2)))) | IN11)) & ((!((((!(IN1)) & (!(IN4))) & (!(IN3))) & IN2)) | IN13)) & ((!(((IN1 & (!(IN4))) & (!(IN3))) & IN2)) | IN14)) & ((!((((!(IN1)) & IN4) & (!(IN3))) & IN2)) | IN15)) & ((!(((IN1 & IN4) & (!(IN3))) & IN2)) | IN16)) & ((!((((!(IN1)) & (!(IN4))) & IN3) & IN2)) | IN17)) & ((!(((IN1 & (!(IN4))) & IN3) & IN2)) | IN18)) & ((!((((!(IN1)) & IN4) & IN3) & IN2)) | IN19)) & ((!(((IN1 & IN4) & IN3) & IN2)) | IN20)

*)

FUNCTION_BLOCK F_CollectInput
  VAR_IN_OUT
      Data : ARRAY[1..20] OF BOOL;
  END_VAR
  VAR_INPUT
      TICK  : BOOL := 0;
      IN1   : BOOL := 0;
      IN2   : BOOL := 0;
      IN3   : BOOL := 0;
      IN4   : BOOL := 0;
      IN5   : BOOL := 0;
      RESET : BOOL := FALSE;
  END_VAR
  VAR_OUTPUT
      Finished : BOOL;
  END_VAR
  VAR
      j    : USINT := 1;
      tock : BOOL  := 0;
  END_VAR
  IF NOT RESET AND tock = NOT TICK THEN
      Data[j]   := IN1;
      Data[j+1] := IN2;
      Data[j+2] := IN3;
      Data[j+3] := IN4;
      Data[j+4] := IN5;
      j := j + 5;
      tock := TICK;
  ELSE
      j := 1;
      tock := 0;
  END_IF;
  Finished := (j > 20);
END_FUNCTION_BLOCK

PROGRAM Boiler
  VAR
    Data  : ARRAY[1..20] OF BOOL;
    Ready : BOOL;
    CollectInput : F_CollectInput;
  END_VAR
  VAR
    TICK     AT %IX1.0 : BOOL;
    IN1      AT %IX0.3 : BOOL;
    IN2      AT %IX0.4 : BOOL;
    IN3      AT %IX0.5 : BOOL;
    IN4      AT %IX0.6 : BOOL;
    IN5      AT %IX0.7 : BOOL;
    OutReady AT %QX0.0 : BOOL := FALSE;
    FeedNext AT %QX0.1 : BOOL := FALSE;
    Out      AT %QX0.2 : BOOL;
  END_VAR
  CollectInput(TICK:=TICK, IN1:=IN1, IN2:=IN2, IN3:=IN3, IN4:=IN4, IN5:=IN5);
  Ready := CollectInput.Finished;
  FeedNext := 1;
  IF Ready THEN
    Out := (((((((((((((((((NOT ((((NOT Data[1]) AND (NOT Data[4])) AND (NOT Data[3])) AND (NOT Data[2]))) OR Data[8]) AND ((NOT (((Data[1] AND (NOT Data[4])) AND (NOT Data[3])) AND (NOT Data[2]))) OR Data[5])) AND ((NOT ((((NOT Data[1]) AND Data[4]) AND (NOT Data[3])) AND (NOT Data[2]))) OR Data[6])) AND ((NOT (((Data[1] AND Data[4]) AND (NOT Data[3])) AND (NOT Data[2]))) OR Data[9])) AND ((NOT ((((NOT Data[1]) AND (NOT Data[4])) AND Data[3]) AND (NOT Data[2]))) OR Data[7])) AND ((NOT (((Data[1] AND (NOT Data[4])) AND Data[3]) AND (NOT Data[2]))) OR Data[10])) AND ((NOT ((((NOT Data[1]) AND Data[4]) AND Data[3]) AND (NOT Data[2]))) OR Data[12])) AND ((NOT (((Data[1] AND Data[4]) AND Data[3]) AND (NOT Data[2]))) OR Data[11])) AND ((NOT ((((NOT Data[1]) AND (NOT Data[4])) AND (NOT Data[3])) AND Data[2])) OR Data[13])) AND ((NOT (((Data[1] AND (NOT Data[4])) AND (NOT Data[3])) AND Data[2])) OR Data[14])) AND ((NOT ((((NOT Data[1]) AND Data[4]) AND (NOT Data[3])) AND Data[2])) OR Data[15])) AND ((NOT (((Data[1] AND Data[4]) AND (NOT Data[3])) AND Data[2])) OR Data[16])) AND ((NOT ((((NOT Data[1]) AND (NOT Data[4])) AND Data[3]) AND Data[2])) OR Data[17])) AND ((NOT (((Data[1] AND (NOT Data[4])) AND Data[3]) AND Data[2])) OR Data[18])) AND ((NOT ((((NOT Data[1]) AND Data[4]) AND Data[3]) AND Data[2])) OR Data[19])) AND ((NOT (((Data[1] AND Data[4]) AND Data[3]) AND Data[2])) OR Data[20]));
    OutReady := 1;
    CollectInput(RESET:=TRUE);
  END_IF;
END_PROGRAM

CONFIGURATION Config0
  RESOURCE Res0 ON PLC
    TASK task0(INTERVAL := T#20ms,PRIORITY := 0);
    PROGRAM instance0 WITH task0 : Boiler;
  END_RESOURCE
END_CONFIGURATION
